(* CODESYS project RobotCell.project

Project tree, tasks and I/O mapping:
  Device : CODESYS Control Win V3 x64, CODESYS, version 3.5.22.40
    application Application
      libraries: Standard, 3.5.22.0 (System); VisuDialogs, * (System)
      task SoftMotion_PlanningTask (freewheeling, priority 15) calls nothing
      task CommTask (cyclic, interval t#50ms, priority 10) calls PRG_Comm
      task MainTask (cyclic, interval 4 ms, priority 1) calls PRG_Main, PRG_Tests, PRG_Recipe_Cell
      task VISU_TASK (cyclic, interval 100 ms, priority 31) calls VisuElems.Visu_Prg, PRG_HMI_Alarms, PRG_HMI_Robot, PRG_HMI_Overview
      axis group AxisGroup_Robot: TRAFO.Kin_ArticulatedRobot_6DOF, axes Axis_J1, Axis_J2, Axis_J3, Axis_J4, Axis_J5, Axis_J6
      Config/
        global variables GVL_Constants
        global variables GVL_CellGeometry
        global variables GVL_Params
        global variables GVL_Config
        global variables GVL_AlarmDefs
      Types/
        data type E_PackMLState
        data type E_PackMLMode
        data type E_PackMLCommand
        data type E_AlarmClass
        data type E_AlarmId
        data type E_Bin
        data type E_Quality
        data type E_DecisionSource
        data type E_PartState
        data type ST_PartRecord
        data type ST_AlarmDef
        data type ST_Alarm
        data type ST_VisionMsg
        data type ST_DecisionMsg
        data type ST_CaptureMsg
        data type E_RobotCmd
        data type E_PickStep
      Interfaces/
        interface I_AlarmSink: Raise, Clear, RaiseEvent
        interface I_Equipment: Reset, HasError, ErrorId
      Framework/
        function block FB_PackMLStateMachine [ST]
        function block FB_AlarmHandler [ST]: Raise, Clear, AcknowledgeAll, GetAlarm, RaiseEvent
        function block FB_PartQueue [ST]: AddRecord, FindIndex, GetRecord, PutRecord, Release, Count, Clear
      Equipment/
        function block FB_PhotoEye [ST]
        function block FB_Bin [ST]: Empty
        function block FB_SafetyMonitor [ST]
        function block FB_VacuumGripper [ST]: Reset, HasError, ErrorId
        function block FB_Conveyor [ST]: Reset, HasError, ErrorId
        function block FB_Robot [ST]: Reset, HasError, ErrorId
        function block FB_JointMonitor [ST]
        function block FB_CameraTrigger [ST]
      Process/
        function F_SelectBin [ST]
        function block FB_PartTracker [ST]: Decide, RaiseAlarm, CurrentX, NextPickable, FindPart, GetRecord, SetState, Count, RaiseEventAlarm, Clear
        function block FB_PickSequence [ST]: Request, NextStep, TrackedPose, GoError
        function block FB_SortingCell [ST]: AlarmState, PlacedCount, RobotMoving, AnyBinFull
      Comm/
        global variables GVL_Bridge
        global variables GVL_Hmi
        function block FB_MessageIntake [ST]
        function block FB_BridgeWatchdog [ST]
      Programs/
        program PRG_Main [ST]
        program PRG_Comm [ST]
      Tests/
        program PRG_TestMotionSmoke [ST]
        program PRG_Tests [ST]
        program PRG_TestTypes [ST]
        program PRG_TestPackML [ST]
        program PRG_TestAlarms [ST]
        program PRG_TestEquipment [ST]
        program PRG_TestMotion [ST]
        program PRG_TestTracking [ST]
        program PRG_TestJointMonitor [ST]
        program PRG_TestPick [ST]
        program PRG_TestCell [ST]
      visualisation Visu_Overview
      data type ST_Recipe_Cell
      global variables GVL_Recipe_Cell
      program PRG_Recipe_Cell [ST]
      Hmi/
        global variables GVL_HmiPanel
        global variables GVL_HmiView
        function block FB_HmiPanel [ST]
        function block FB_HmiView [ST]
      program PRG_HMI_Alarms [ST]
      visualisation Visu_Robot
      image pool IP_Robot
      program PRG_HMI_Robot [ST]
      program PRG_HMI_Overview [ST]
      image pool IP_Overview
      visualisation Visu_Alarms
      image pool IP_Alarms
    SoftMotion General Axis Pool : SoftMotion General Axis Pool, CODESYS, version 4.11.0.0
      Axis_J1 : SM_Drive_Virtual, CODESYS, order no. 1805, version 4.18.0.0
          settings: wDriveID = 0; fSWMaxVelocity = 180; fSWLimitPositive = 170; fSWLimitNegative = -170; bSWLimitEnable = true
      Axis_J2 : SM_Drive_Virtual, CODESYS, order no. 1805, version 4.18.0.0
          settings: fSWMaxVelocity = 180; fSWLimitPositive = 150; fSWLimitNegative = -90; bSWLimitEnable = true
      Axis_J3 : SM_Drive_Virtual, CODESYS, order no. 1805, version 4.18.0.0
          settings: wDriveID = 2; fSWMaxVelocity = 180; fSWLimitPositive = 150; fSWLimitNegative = -120; bSWLimitEnable = true
      Axis_J4 : SM_Drive_Virtual, CODESYS, order no. 1805, version 4.18.0.0
          settings: wDriveID = 3; fSWMaxVelocity = 360; fSWLimitPositive = 180; fSWLimitNegative = -180; bSWLimitEnable = true
      Axis_J5 : SM_Drive_Virtual, CODESYS, order no. 1805, version 4.18.0.0
          settings: wDriveID = 4; fSWMaxVelocity = 360; fSWLimitPositive = 120; fSWLimitNegative = -120; bSWLimitEnable = true
      Axis_J6 : SM_Drive_Virtual, CODESYS, order no. 1805, version 4.18.0.0
          settings: wDriveID = 5; fSWMaxVelocity = 360; fSWLimitPositive = 360; fSWLimitNegative = -360; bSWLimitEnable = true
      Axis_Conveyor : SM_Drive_Virtual, CODESYS, order no. 1805, version 4.18.0.0
          settings: wDriveID = 6; fSWMaxVelocity = 400; bSWLimitEnable = false
  libraries: VisuSymbols, 4.5.0.0 (System)
  5ce3da45-db07-42e7-a21c-a00fff4ed8f6|C:\Users\AvazA\AppData\Local\Temp\cmcp-visu-UXzo4K\ic_alarm_24_80868c.svg
  5ce3da45-db07-42e7-a21c-a00fff4ed8f6|C:\Users\AvazA\AppData\Local\Temp\cmcp-visu-UXzo4K\ic_check_27_1a232d.svg
  5ce3da45-db07-42e7-a21c-a00fff4ed8f6|C:\Users\AvazA\AppData\Local\Temp\cmcp-visu-UXzo4K\ic_pause_27_1a232d.svg
  5ce3da45-db07-42e7-a21c-a00fff4ed8f6|C:\Users\AvazA\AppData\Local\Temp\cmcp-visu-UXzo4K\ic_play_27_1a232d.svg
  5ce3da45-db07-42e7-a21c-a00fff4ed8f6|C:\Users\AvazA\AppData\Local\Temp\cmcp-visu-UXzo4K\stn_bin_on_48x48.svg
  5ce3da45-db07-42e7-a21c-a00fff4ed8f6|C:\Users\AvazA\AppData\Local\Temp\cmcp-visu-vSJax5\ic_stop_30_66727e.svg
  5ce3da45-db07-42e7-a21c-a00fff4ed8f6|C:\Users\AvazA\AppData\Local\Temp\cmcp-visu-vSJax5\ic_fault_30_d72332.svg
  5ce3da45-db07-42e7-a21c-a00fff4ed8f6|C:\Users\AvazA\AppData\Local\Temp\cmcp-visu-vSJax5\ic_pause_30_ffbb00.svg
  5ce3da45-db07-42e7-a21c-a00fff4ed8f6|C:\Users\AvazA\AppData\Local\Temp\cmcp-visu-vSJax5\ic_warning_30_ffbb00.svg
  5ce3da45-db07-42e7-a21c-a00fff4ed8f6|C:\Users\AvazA\AppData\Local\Temp\cmcp-visu-vSJax5\ic_manual_30_2f5d8a.svg
  5ce3da45-db07-42e7-a21c-a00fff4ed8f6|C:\Users\AvazA\AppData\Local\Temp\cmcp-visu-vSJax5\ic_play_30_66727e.svg
  5ce3da45-db07-42e7-a21c-a00fff4ed8f6|C:\Users\AvazA\AppData\Local\Temp\cmcp-visu-vSJax5\ic_login_27_1a232d.svg
  5ce3da45-db07-42e7-a21c-a00fff4ed8f6|C:\Users\AvazA\AppData\Local\Temp\cmcp-visu-vSJax5\ic_reset_27_1a232d.svg
  5ce3da45-db07-42e7-a21c-a00fff4ed8f6|C:\Users\AvazA\AppData\Local\Temp\cmcp-visu-vSJax5\ic_play_27_ffffff.svg
  5ce3da45-db07-42e7-a21c-a00fff4ed8f6|C:\Users\AvazA\AppData\Local\Temp\cmcp-visu-UXzo4K\sign_warning_30.svg
  5ce3da45-db07-42e7-a21c-a00fff4ed8f6|C:\Users\AvazA\AppData\Local\Temp\cmcp-visu-UXzo4K\ic_speed_24_80868c.svg
  5ce3da45-db07-42e7-a21c-a00fff4ed8f6|C:\Users\AvazA\AppData\Local\Temp\cmcp-visu-UXzo4K\ic_warning_30_ffbb00.svg
  5ce3da45-db07-42e7-a21c-a00fff4ed8f6|C:\Users\AvazA\AppData\Local\Temp\cmcp-visu-UXzo4K\ic_pause_30_ffbb00.svg
  5ce3da45-db07-42e7-a21c-a00fff4ed8f6|C:\Users\AvazA\AppData\Local\Temp\cmcp-visu-UXzo4K\ic_fault_30_d72332.svg
  5ce3da45-db07-42e7-a21c-a00fff4ed8f6|C:\Users\AvazA\AppData\Local\Temp\cmcp-visu-UXzo4K\ic_count_24_80868c.svg
  5ce3da45-db07-42e7-a21c-a00fff4ed8f6|C:\Users\AvazA\AppData\Local\Temp\cmcp-visu-UXzo4K\stn_bin_off_48x48.svg
  text list GlobalTextList
  5ce3da45-db07-42e7-a21c-a00fff4ed8f6|C:\Users\AvazA\AppData\Local\Temp\cmcp-visu-vSJax5\ic_stop_27_1a232d.svg
  5ce3da45-db07-42e7-a21c-a00fff4ed8f6|C:\Users\AvazA\AppData\Local\Temp\cmcp-visu-vSJax5\ic_home_33_5c636a.svg
  5ce3da45-db07-42e7-a21c-a00fff4ed8f6|C:\Users\AvazA\AppData\Local\Temp\cmcp-visu-vSJax5\ic_machine_33_2f5d8a.svg
  5ce3da45-db07-42e7-a21c-a00fff4ed8f6|C:\Users\AvazA\AppData\Local\Temp\cmcp-visu-vSJax5\ic_alarm_33_5c636a.svg
  5ce3da45-db07-42e7-a21c-a00fff4ed8f6|C:\Users\AvazA\AppData\Local\Temp\cmcp-visu-vSJax5\ic_manual_24_80868c.svg
  5ce3da45-db07-42e7-a21c-a00fff4ed8f6|C:\Users\AvazA\AppData\Local\Temp\cmcp-visu-vSJax5\ic_info_24_80868c.svg
  5ce3da45-db07-42e7-a21c-a00fff4ed8f6|C:\Users\AvazA\AppData\Local\Temp\cmcp-visu-vSJax5\ic_speed_24_80868c.svg
  5ce3da45-db07-42e7-a21c-a00fff4ed8f6|C:\Users\AvazA\AppData\Local\Temp\cmcp-visu-vSJax5\ic_machine_24_80868c.svg
  5ce3da45-db07-42e7-a21c-a00fff4ed8f6|C:\Users\AvazA\AppData\Local\Temp\cmcp-visu-UXzo4K\stn_robot6_off_48x48.svg
  5ce3da45-db07-42e7-a21c-a00fff4ed8f6|C:\Users\AvazA\AppData\Local\Temp\cmcp-visu-UXzo4K\ic_manual_23_2f5d8a.svg
  5ce3da45-db07-42e7-a21c-a00fff4ed8f6|C:\Users\AvazA\AppData\Local\Temp\cmcp-visu-UXzo4K\stn_camera_on_48x48.svg
  5ce3da45-db07-42e7-a21c-a00fff4ed8f6|C:\Users\AvazA\AppData\Local\Temp\cmcp-visu-UXzo4K\stn_camera_off_48x48.svg
  5ce3da45-db07-42e7-a21c-a00fff4ed8f6|C:\Users\AvazA\AppData\Local\Temp\cmcp-visu-UXzo4K\sign_alarm_27.svg
  5ce3da45-db07-42e7-a21c-a00fff4ed8f6|C:\Users\AvazA\AppData\Local\Temp\cmcp-visu-UXzo4K\stn_conveyor_on_48x14.svg
  5ce3da45-db07-42e7-a21c-a00fff4ed8f6|C:\Users\AvazA\AppData\Local\Temp\cmcp-visu-UXzo4K\stn_conveyor_off_48x14.svg
  5ce3da45-db07-42e7-a21c-a00fff4ed8f6|C:\Users\AvazA\AppData\Local\Temp\cmcp-visu-UXzo4K\sign_stop_13.svg
  5ce3da45-db07-42e7-a21c-a00fff4ed8f6|C:\Users\AvazA\AppData\Local\Temp\cmcp-visu-UXzo4K\sign_run_15.svg
  5ce3da45-db07-42e7-a21c-a00fff4ed8f6|C:\Users\AvazA\AppData\Local\Temp\cmcp-visu-UXzo4K\arrow_r_15_92979b.svg
  5ce3da45-db07-42e7-a21c-a00fff4ed8f6|C:\Users\AvazA\AppData\Local\Temp\cmcp-visu-UXzo4K\ic_alarm_33_5c636a.svg
  5ce3da45-db07-42e7-a21c-a00fff4ed8f6|C:\Users\AvazA\AppData\Local\Temp\cmcp-visu-UXzo4K\ic_machine_33_5c636a.svg
  5ce3da45-db07-42e7-a21c-a00fff4ed8f6|C:\Users\AvazA\AppData\Local\Temp\cmcp-visu-UXzo4K\ic_home_33_2f5d8a.svg
  5ce3da45-db07-42e7-a21c-a00fff4ed8f6|C:\Users\AvazA\AppData\Local\Temp\cmcp-visu-UXzo4K\ic_stop_27_1a232d.svg
  5ce3da45-db07-42e7-a21c-a00fff4ed8f6|C:\Users\AvazA\AppData\Local\Temp\cmcp-visu-UXzo4K\ic_play_27_ffffff.svg
  5ce3da45-db07-42e7-a21c-a00fff4ed8f6|C:\Users\AvazA\AppData\Local\Temp\cmcp-visu-UXzo4K\ic_reset_27_1a232d.svg
  5ce3da45-db07-42e7-a21c-a00fff4ed8f6|C:\Users\AvazA\AppData\Local\Temp\cmcp-visu-UXzo4K\ic_login_27_1a232d.svg
  5ce3da45-db07-42e7-a21c-a00fff4ed8f6|C:\Users\AvazA\AppData\Local\Temp\cmcp-visu-UXzo4K\ic_play_30_66727e.svg
  5ce3da45-db07-42e7-a21c-a00fff4ed8f6|C:\Users\AvazA\AppData\Local\Temp\cmcp-visu-UXzo4K\ic_manual_30_2f5d8a.svg
  5ce3da45-db07-42e7-a21c-a00fff4ed8f6|C:\Users\AvazA\AppData\Local\Temp\cmcp-visu-UXzo4K\ic_stop_30_66727e.svg
  5ce3da45-db07-42e7-a21c-a00fff4ed8f6|C:\Users\AvazA\AppData\Local\Temp\cmcp-visu-UXzo4K\stn_robot6_on_48x48.svg
  5ce3da45-db07-42e7-a21c-a00fff4ed8f6|C:\Users\AvazA\AppData\Local\Temp\cmcp-visu-UXzo4K\stn_gripper_on_48x48.svg
  5ce3da45-db07-42e7-a21c-a00fff4ed8f6|C:\Users\AvazA\AppData\Local\Temp\cmcp-visu-UXzo4K\stn_gripper_off_48x48.svg
  5ce3da45-db07-42e7-a21c-a00fff4ed8f6|C:\Users\AvazA\AppData\Local\Temp\cmcp-visu-6UqmBO\ic_check_27_1a232d.svg
  5ce3da45-db07-42e7-a21c-a00fff4ed8f6|C:\Users\AvazA\AppData\Local\Temp\cmcp-visu-6UqmBO\ic_warning_24_80868c.svg
  5ce3da45-db07-42e7-a21c-a00fff4ed8f6|C:\Users\AvazA\AppData\Local\Temp\cmcp-visu-6UqmBO\ic_alarm_24_80868c.svg
  5ce3da45-db07-42e7-a21c-a00fff4ed8f6|C:\Users\AvazA\AppData\Local\Temp\cmcp-visu-6UqmBO\ic_alarm_33_2f5d8a.svg
  5ce3da45-db07-42e7-a21c-a00fff4ed8f6|C:\Users\AvazA\AppData\Local\Temp\cmcp-visu-6UqmBO\ic_machine_33_5c636a.svg
  5ce3da45-db07-42e7-a21c-a00fff4ed8f6|C:\Users\AvazA\AppData\Local\Temp\cmcp-visu-6UqmBO\ic_home_33_5c636a.svg
  5ce3da45-db07-42e7-a21c-a00fff4ed8f6|C:\Users\AvazA\AppData\Local\Temp\cmcp-visu-6UqmBO\ic_stop_27_1a232d.svg
  5ce3da45-db07-42e7-a21c-a00fff4ed8f6|C:\Users\AvazA\AppData\Local\Temp\cmcp-visu-6UqmBO\ic_play_27_ffffff.svg
  5ce3da45-db07-42e7-a21c-a00fff4ed8f6|C:\Users\AvazA\AppData\Local\Temp\cmcp-visu-6UqmBO\ic_reset_27_1a232d.svg
  5ce3da45-db07-42e7-a21c-a00fff4ed8f6|C:\Users\AvazA\AppData\Local\Temp\cmcp-visu-6UqmBO\ic_login_27_1a232d.svg
  5ce3da45-db07-42e7-a21c-a00fff4ed8f6|C:\Users\AvazA\AppData\Local\Temp\cmcp-visu-6UqmBO\ic_play_30_66727e.svg
  5ce3da45-db07-42e7-a21c-a00fff4ed8f6|C:\Users\AvazA\AppData\Local\Temp\cmcp-visu-6UqmBO\ic_manual_30_2f5d8a.svg
  5ce3da45-db07-42e7-a21c-a00fff4ed8f6|C:\Users\AvazA\AppData\Local\Temp\cmcp-visu-6UqmBO\ic_warning_30_ffbb00.svg
  5ce3da45-db07-42e7-a21c-a00fff4ed8f6|C:\Users\AvazA\AppData\Local\Temp\cmcp-visu-6UqmBO\ic_pause_30_ffbb00.svg
  5ce3da45-db07-42e7-a21c-a00fff4ed8f6|C:\Users\AvazA\AppData\Local\Temp\cmcp-visu-6UqmBO\ic_fault_30_d72332.svg
  5ce3da45-db07-42e7-a21c-a00fff4ed8f6|C:\Users\AvazA\AppData\Local\Temp\cmcp-visu-6UqmBO\ic_stop_30_66727e.svg
  5ce3da45-db07-42e7-a21c-a00fff4ed8f6|C:\Users\AvazA\AppData\Local\Temp\cmcp-visu-UXzo4K\ic_info_24_80868c.svg
*)

// Device/Application/Types/E_PackMLState
// PackML unit states, numbered as in ISA-TR88.00.02.
{attribute 'qualified_only'}
{attribute 'strict'}
TYPE E_PackMLState :
(
    Undefined := 0,
    Clearing := 1,
    Stopped := 2,
    Starting := 3,
    Idle := 4,
    Suspended := 5,
    Execute := 6,
    Stopping := 7,
    Aborting := 8,
    Aborted := 9,
    Holding := 10,
    Held := 11,
    Unholding := 12,
    Suspending := 13,
    Unsuspending := 14,
    Resetting := 15,
    Completing := 16,
    Complete := 17
);
END_TYPE

// Device/Application/Types/E_PackMLMode
// PackML unit modes used by this cell.
{attribute 'qualified_only'}
{attribute 'strict'}
TYPE E_PackMLMode :
(
    Production := 1,
    Maintenance := 2,
    Manual := 3
);
END_TYPE

// Device/Application/Types/E_PackMLCommand
// PackML state commands.
{attribute 'qualified_only'}
{attribute 'strict'}
TYPE E_PackMLCommand :
(
    None := 0,
    Reset := 1,
    Start := 2,
    Stop := 3,
    Hold := 4,
    Unhold := 5,
    Suspend := 6,
    Unsuspend := 7,
    Abort := 8,
    Clear := 9,
    Complete := 10
);
END_TYPE

// Device/Application/Types/E_AlarmClass
// Alarm classes (ISA-18.2 style priorities). Critical -> Abort, Error -> Stop.
{attribute 'qualified_only'}
{attribute 'strict'}
TYPE E_AlarmClass :
(
    Info := 0,
    Warning := 1,
    Error := 2,
    Critical := 3
);
END_TYPE

// Device/Application/Types/E_AlarmId
// Every alarm of the cell. Definitions (class, text) are in GVL_AlarmDefs.
{attribute 'qualified_only'}
{attribute 'strict'}
TYPE E_AlarmId :
(
    None := 0,
    EStop := 1,
    DoorOpen := 2,
    BridgeLost := 3,
    AxisGroupError := 4,
    ConveyorError := 5,
    FollowingErrorWarn := 6,
    FollowingErrorFault := 7,
    FeedbackStale := 8,
    VacuumNoGrip := 9,
    VacuumLost := 10,
    PartMissed := 11,
    BinFull := 12,
    VisionMissing := 13,
    DecisionFallback := 14,
    LowConfidence := 15,
    QueueOverflow := 16
);
END_TYPE

// Device/Application/Types/E_Bin
// Output bins: one per good part type, then the quality bins.
{attribute 'qualified_only'}
{attribute 'strict'}
TYPE E_Bin :
(
    TypeA := 0,
    TypeB := 1,
    TypeC := 2,
    Rework := 3,
    Scrap := 4,
    Quarantine := 5
);
END_TYPE

// Device/Application/Types/E_Quality
// Quality disposition of a part (spec section 6.3).
{attribute 'qualified_only'}
{attribute 'strict'}
TYPE E_Quality :
(
    Unknown := 0,
    Ok := 1,
    Rework := 2,
    Scrap := 3
);
END_TYPE

// Device/Application/Types/E_DecisionSource
// Where a part's quality decision came from.
{attribute 'qualified_only'}
{attribute 'strict'}
TYPE E_DecisionSource :
(
    None := 0,
    Ai := 1,
    Fallback := 2
);
END_TYPE

// Device/Application/Types/E_PartState
// Life cycle of a tracked part.
{attribute 'qualified_only'}
{attribute 'strict'}
TYPE E_PartState :
(
    Free := 0,
    Captured := 1,
    Identified := 2,
    Decided := 3,
    Scheduled := 4,
    Picked := 5,
    Placed := 6,
    Missed := 7,
    Dropped := 8
);
END_TYPE

// Device/Application/Types/ST_PartRecord
// One tracked part. Positions are in the belt frame at capture time (mm, degrees).
TYPE ST_PartRecord :
STRUCT
    udiPartId : UDINT;
    lrBeltPosAtCapture : LREAL;         // conveyor axis position when PE1 triggered [mm]
    xVisionValid : BOOL;
    usiClass : USINT;                   // detector class index 0..2
    rConfidence : REAL;                 // detector confidence 0..1
    lrX : LREAL;                        // belt frame X at capture [mm]
    lrY : LREAL;                        // belt frame Y [mm]
    lrTheta : LREAL;                    // orientation about Z [deg]
    eQuality : E_Quality;
    rQualityProb : REAL;                // probability of the chosen quality option
    xIdentReliable : BOOL;
    eDecisionSource : E_DecisionSource;
    eTargetBin : E_Bin;
    eState : E_PartState;
    tCaptured : TIME;                   // TIME() at capture
END_STRUCT
END_TYPE

// Device/Application/Types/ST_AlarmDef
// Static definition of one alarm.
TYPE ST_AlarmDef :
STRUCT
    eClass : E_AlarmClass;
    sText : STRING(80);
END_STRUCT
END_TYPE

// Device/Application/Types/ST_Alarm
// Runtime state of one alarm.
TYPE ST_Alarm :
STRUCT
    eClass : E_AlarmClass;
    xActive : BOOL;
    xAcked : BOOL := TRUE;              // no pending acknowledgement
    tRaised : TIME;
END_STRUCT
END_TYPE

// Device/Application/Types/ST_VisionMsg
// Vision result written by the bridge. A new message has a new udiSeq.
TYPE ST_VisionMsg :
STRUCT
    udiSeq : UDINT;
    udiPartId : UDINT;
    xValid : BOOL;
    usiClass : USINT;
    rConfidence : REAL;
    lrX : LREAL;                        // belt frame [mm]
    lrY : LREAL;                        // belt frame [mm]
    lrTheta : LREAL;                    // [deg]
END_STRUCT
END_TYPE

// Device/Application/Types/ST_DecisionMsg
// Quality decision written by the bridge (THX-02). A new message has a new udiSeq.
TYPE ST_DecisionMsg :
STRUCT
    udiSeq : UDINT;
    udiPartId : UDINT;
    eQuality : E_Quality;
    rQualityProb : REAL;
    xIdentReliable : BOOL;
END_STRUCT
END_TYPE

// Device/Application/Types/ST_CaptureMsg
// Capture request from the PLC to the bridge. A new request has a new udiSeq.
TYPE ST_CaptureMsg :
STRUCT
    udiSeq : UDINT;
    udiPartId : UDINT;
    lrBeltPos : LREAL;                  // conveyor axis position at the trigger [mm]
END_STRUCT
END_TYPE

// Device/Application/Types/E_RobotCmd
// Commands of FB_Robot (start on a rising edge of xExecute).
{attribute 'qualified_only'}
{attribute 'strict'}
TYPE E_RobotCmd :
(
    None := 0,
    MovePtpAcs := 1,       // point-to-point, target in joint space
    MoveLinMcs := 2,       // linear, target in machine coordinates
    MoveLinPcs1 := 3,      // linear, target in PCS_1 (conveyor tracking frame)
    Stop := 4,             // controlled stop, aborts any motion
    Reset := 5,            // reset axis group errors
    MovePtpMcs := 6        // point-to-point, Cartesian target in machine coordinates
);
END_TYPE

// Device/Application/Types/E_PickStep
// Steps of FB_PickSequence.
{attribute 'qualified_only'}
{attribute 'strict'}
TYPE E_PickStep :
(
    Idle := 0,
    MoveHome := 1,
    MoveReady := 2,
    WaitPart := 3,
    StartTracking := 4,
    Approach := 5,
    Descend := 6,
    Grip := 7,
    Lift := 8,
    MoveToBin := 9,
    Release := 10,
    Retract := 11,
    Aborting := 12,
    Aborted := 13,
    Error := 14,
    RecoverLift := 15       // after an abort with a part on the cup: straight up first
);
END_TYPE

// Device/Application/ST_Recipe_Cell
TYPE ST_Recipe_Cell :
STRUCT
    lrBeltSpeed : LREAL; // GVL_Params.lrBeltSpeed
    lrApproachHeight : LREAL; // GVL_Params.lrApproachHeight
    lrPickDepth : LREAL; // GVL_Params.lrPickDepth
    lrLinVelocity : LREAL; // GVL_Params.lrLinVelocity
    lrLinAccel : LREAL; // GVL_Params.lrLinAccel
    lrLinJerk : LREAL; // GVL_Params.lrLinJerk
    lrPtpVelFactor : LREAL; // GVL_Params.lrPtpVelFactor
    rConfidenceThreshold : REAL; // GVL_Params.rConfidenceThreshold
    tDecisionDeadline : TIME; // GVL_Params.tDecisionDeadline
    tVacuumTimeout : TIME; // GVL_Params.tVacuumTimeout
    lrFollowErrWarn : LREAL; // GVL_Params.lrFollowErrWarn
    lrFollowErrFault : LREAL; // GVL_Params.lrFollowErrFault
    tFeedbackTimeout : TIME; // GVL_Params.tFeedbackTimeout
END_STRUCT
END_TYPE

// Device/Application/Config/GVL_Constants
// Project-wide constants. Values that change per recipe live in GVL_Params, not here.
{attribute 'qualified_only'}
VAR_GLOBAL CONSTANT
    PROJECT_VERSION : STRING := '0.7.0';
END_VAR

// Device/Application/Config/GVL_CellGeometry
// Fixed geometry of the cell. Units: mm and degrees, robot base frame (Z up).
// Kinematics values must match the axis group AxisGroup_Robot (plc/scripts/build_softmotion_base.py).
// Orientations (A, B, C): B = 180 points the tool straight down (verified in simulation).
{attribute 'qualified_only'}
VAR_GLOBAL CONSTANT
    // Kin_ArticulatedRobot_6DOF parameters [mm]
    ROBOT_A1 : LREAL := 50;
    ROBOT_D1 : LREAL := 400;
    ROBOT_A2 : LREAL := 450;
    ROBOT_A3 : LREAL := 50;
    ROBOT_D3 : LREAL := 0;
    ROBOT_D4 : LREAL := 450;
    ROBOT_D6 : LREAL := 120;                 // flange + suction tool

    // Tool pointing straight down
    TOOL_DOWN_A : LREAL := 0;
    TOOL_DOWN_B : LREAL := 180;
    TOOL_DOWN_C : LREAL := 180;

    // Conveyor belt frame: origin at the infeed, +X along the flow direction.
    BELT_ORIGIN : MC_COORD_REF := (X := -1500, Y := -550, Z := 0, A := 0, B := 0, C := 0);
    BELT_SURFACE_Z : LREAL := 0;
    PE1_X : LREAL := 300;                    // camera trigger photo-eye, belt frame [mm]
    PE2_X : LREAL := 1050;                   // pick window start, belt frame [mm]
    PICK_WINDOW_END_X : LREAL := 1750;       // pick window end, belt frame [mm]
    PICK_MARGIN : LREAL := 300;              // do not start a pick this close to the window end [mm]
    // Grip height of each part class above the belt [mm]: the top surface under the suction
    // cup (config/parts.yaml classes, tools/fetch_objects.py meta.json; a unit test keeps
    // both equal)
    PART_HEIGHTS : ARRAY[0..2] OF LREAL := [56.39, 81.19, 83.46];

    // Home position, joint space [deg]
    HOME_ACS : SMC_POS_REF := (a := (a0 := 0, a1 := -30, a2 := 60, a3 := 0, a4 := 60, a5 := 0));
    // Waiting pose above the pick window, tool down (machine coordinates)
    READY_POSE : MC_COORD_REF := (X := -100, Y := -550, Z := 300, A := 0, B := 180, C := 180);
    RETRACT_HEIGHT : LREAL := 100;           // lift above the bin drop pose after release [mm]

    // Drop poses above the bins (tool pointing down), machine coordinates [mm, deg]. Z 300: a
    // held part up to 90 mm tall clears the 160 mm bin rim by 50 mm.
    BIN_DROP : ARRAY[E_Bin.TypeA..E_Bin.Quarantine] OF MC_COORD_REF := [
        (X := -500, Y := 550, Z := 300, A := 0, B := 180, C := 180),
        (X := -300, Y := 550, Z := 300, A := 0, B := 180, C := 180),
        (X := -100, Y := 550, Z := 300, A := 0, B := 180, C := 180),
        (X := 100, Y := 550, Z := 300, A := 0, B := 180, C := 180),
        (X := 300, Y := 550, Z := 300, A := 0, B := 180, C := 180),
        (X := 500, Y := 550, Z := 300, A := 0, B := 180, C := 180)];
END_VAR

// Device/Application/Config/GVL_Params
// Process parameters. Retained; written by the recipes (Standard / HighSpeed).
{attribute 'qualified_only'}
VAR_GLOBAL RETAIN
    lrBeltSpeed : LREAL := 100;              // conveyor speed [mm/s]
    lrApproachHeight : LREAL := 80;          // approach / lift height above the part [mm]
    lrPickDepth : LREAL := 5;                // how far below the part top the cup goes [mm]
    lrLinVelocity : LREAL := 500;            // linear path velocity [mm/s]
    lrLinAccel : LREAL := 2000;              // linear path acceleration [mm/s2]
    lrLinJerk : LREAL := 20000;              // linear path jerk [mm/s3]
    lrPtpVelFactor : LREAL := 0.5;           // PTP velocity factor ]0, 1]
    rConfidenceThreshold : REAL := 0.6;      // below this the part goes to quarantine
    tDecisionDeadline : TIME := T#2S500MS;   // fallback if no decision by then
    tVacuumTimeout : TIME := T#500MS;        // no grip -> error
    lrFollowErrWarn : LREAL := 2.0;          // following error warning [deg]
    lrFollowErrFault : LREAL := 5.0;         // following error fault [deg]
    tFeedbackTimeout : TIME := T#500MS;      // joint feedback must update within this time
    aClassToBin : ARRAY[0..2] OF E_Bin := [E_Bin.TypeA, E_Bin.TypeB, E_Bin.TypeC];
END_VAR

// Device/Application/Config/GVL_Config
// Build/run configuration.
{attribute 'qualified_only'}
VAR_GLOBAL
    // Joint feedback := setpoint (no staleness check) unless the twin reports itself active through
    // GVL_Bridge.xTwinActive. FALSE forces real feedback even without the twin.
    xFeedbackLoopback : BOOL := TRUE;
    // The sorting cell runs in PRG_Main. Simulation tests of single blocks switch it off so their
    // harnesses can own the robot and the conveyor.
    xCellEnabled : BOOL := TRUE;
END_VAR
VAR_GLOBAL CONSTANT
    MAX_PARTS : UINT := 32;                  // capacity of the part queue
END_VAR

// Device/Application/Config/GVL_AlarmDefs
// Alarm definitions: class and operator text for every E_AlarmId.
// Critical -> PackML Abort, Error -> Stop, Warning -> no state change (BinFull suspends the unit).
{attribute 'qualified_only'}
VAR_GLOBAL CONSTANT
    aDefs : ARRAY[E_AlarmId.None..E_AlarmId.QueueOverflow] OF ST_AlarmDef := [
        (eClass := E_AlarmClass.Info, sText := 'No alarm'),
        (eClass := E_AlarmClass.Critical, sText := 'Emergency stop pressed'),
        (eClass := E_AlarmClass.Critical, sText := 'Safety door opened in automatic mode'),
        (eClass := E_AlarmClass.Critical, sText := 'Connection to the digital twin bridge lost'),
        (eClass := E_AlarmClass.Critical, sText := 'Robot axis group error'),
        (eClass := E_AlarmClass.Error, sText := 'Conveyor axis error'),
        (eClass := E_AlarmClass.Warning, sText := 'Joint following error above warning limit'),
        (eClass := E_AlarmClass.Critical, sText := 'Joint following error above fault limit'),
        (eClass := E_AlarmClass.Critical, sText := 'Joint feedback not updated'),
        (eClass := E_AlarmClass.Error, sText := 'Vacuum not reached - part not gripped'),
        (eClass := E_AlarmClass.Error, sText := 'Vacuum lost while carrying a part'),
        (eClass := E_AlarmClass.Warning, sText := 'Part left the pick window unpicked'),
        (eClass := E_AlarmClass.Warning, sText := 'A bin is full - cell suspended until it is emptied'),
        (eClass := E_AlarmClass.Warning, sText := 'No vision result for a captured part'),
        (eClass := E_AlarmClass.Warning, sText := 'AI decision late - fallback rule used'),
        (eClass := E_AlarmClass.Warning, sText := 'Low detection confidence - part quarantined'),
        (eClass := E_AlarmClass.Error, sText := 'Part queue full')];
END_VAR

// Device/Application/Comm/GVL_Bridge
// Exchange with the Python bridge over OPC UA (published by the symbol configuration).
// Tag names for the bridge: config/opcua_tags.yaml. In Phase 1, tests write the inputs.
{attribute 'qualified_only'}
{attribute 'symbol' := 'readwrite'}
VAR_GLOBAL
    // --- inputs (bridge -> PLC) ---
    xHeartbeat : BOOL;                                     // toggled by the bridge every cycle
    xTwinActive : BOOL;                                    // the twin delivers joint feedback
    aJointPosFb : ARRAY[1..6] OF LREAL;                    // measured joint positions [deg]
    aJointTorqueFb : ARRAY[1..6] OF LREAL;                 // measured joint torques [Nm]
    udiFeedbackSeq : UDINT;                                // increments with every feedback sample
    udiFeedbackForSeq : UDINT;                             // udiSetpointSeq the feedback belongs to
    xPE1 : BOOL;                                           // photo-eye at the camera
    xPE2 : BOOL;                                           // photo-eye at the pick window start
    xVacuumOk : BOOL;                                      // vacuum switch of the suction cup
    axBinFull : ARRAY[E_Bin.TypeA..E_Bin.Quarantine] OF BOOL;
    xDoorClosed : BOOL := TRUE;                            // safety door (TRUE = closed)
    xEStopOk : BOOL := TRUE;                               // emergency stop circuit (TRUE = not pressed)
    stVision : ST_VisionMsg;
    stDecision : ST_DecisionMsg;
    xDecisionActive : BOOL;                                // an AI decision service answers stDecision
    // --- outputs (PLC -> bridge) ---
    aJointPosSp : ARRAY[1..6] OF LREAL;                    // joint setpoints [deg]
    udiSetpointSeq : UDINT;                                // increments with every setpoint sample
    lrBeltPos : LREAL;                                     // conveyor position [mm]
    lrBeltVel : LREAL;                                     // conveyor velocity [mm/s]
    xVacuumOn : BOOL;                                      // vacuum valve
    stCapture : ST_CaptureMsg;
    eState : E_PackMLState;
    eMode : E_PackMLMode;
    // --- diagnostics (PLC -> bridge, HMI) ---
    eNewestAlarm : E_AlarmId;
    xAlarmError : BOOL;                                    // an Error-class alarm is active
    xAlarmCritical : BOOL;                                 // a Critical-class alarm is active
    ePickStep : E_PickStep;
    iWorstJoint : INT;                                     // joint with the largest following error
    aFollowingError : ARRAY[1..6] OF LREAL;                // [deg]
END_VAR

// Device/Application/Comm/GVL_Hmi
// Operator commands from the HMI (CODESYS Visualization) and, for tests and the HMI of later
// phases, over OPC UA (published by the symbol configuration).
{attribute 'qualified_only'}
{attribute 'symbol' := 'readwrite'}
VAR_GLOBAL
    eCommand : E_PackMLCommand;
    eModeRequest : E_PackMLMode := E_PackMLMode.Production;
    xAlarmAck : BOOL;
    axJogPlus : ARRAY[1..6] OF BOOL;
    axJogMinus : ARRAY[1..6] OF BOOL;
    rOverride : REAL := 1.0;                               // speed override ]0, 1]
END_VAR

// Device/Application/GVL_Recipe_Cell
// Recipes 'Cell', generated by codesys-mcp-toolkit (create_recipes). RETAIN: values saved from the HMI survive a power cycle.
VAR_GLOBAL RETAIN
    aRecipes : ARRAY[0..1] OF ST_Recipe_Cell := [(lrBeltSpeed := 100.0, lrApproachHeight := 80.0, lrPickDepth := 5.0, lrLinVelocity := 500.0, lrLinAccel := 2000.0, lrLinJerk := 20000.0, lrPtpVelFactor := 0.5, rConfidenceThreshold := 0.6, tDecisionDeadline := T#2S500MS, tVacuumTimeout := T#500MS, lrFollowErrWarn := 2.0, lrFollowErrFault := 5.0, tFeedbackTimeout := T#500MS), (lrBeltSpeed := 200.0, lrApproachHeight := 80.0, lrPickDepth := 5.0, lrLinVelocity := 800.0, lrLinAccel := 3000.0, lrLinJerk := 20000.0, lrPtpVelFactor := 0.8, rConfidenceThreshold := 0.6, tDecisionDeadline := T#2S500MS, tVacuumTimeout := T#500MS, lrFollowErrWarn := 2.0, lrFollowErrFault := 5.0, tFeedbackTimeout := T#500MS)];
END_VAR
VAR_GLOBAL CONSTANT
    asNames : ARRAY[0..1] OF STRING(32) := ['Standard', 'HighSpeed'];
    iCount : INT := 2;
END_VAR

// Device/Application/Hmi/GVL_HmiPanel
// Operator panel of the CODESYS Visualization: buttons and selectors write here; FB_HmiPanel
// turns them into the cell's commands (GVL_Hmi). Buttons are one-shot: cleared after use.
{attribute 'qualified_only'}
VAR_GLOBAL
    xStart : BOOL;
    xStop : BOOL;
    xReset : BOOL;
    xClear : BOOL;
    xAbort : BOOL;
    xSuspend : BOOL;
    xUnsuspend : BOOL;
    xAckAll : BOOL;                                        // acknowledge all alarms
    iModeSelect : INT := 1;                                // 1 Production, 2 Maintenance, 3 Manual
END_VAR

// Device/Application/Hmi/GVL_HmiView
// Display data for the CODESYS Visualization, prepared by FB_HmiView (no logic in screens).
{attribute 'qualified_only'}
VAR_GLOBAL
    sState : STRING(20);                                   // PackML state
    sMode : STRING(20);                                    // PackML mode
    sPickStep : STRING(20);                                // robot sequence step
    sNewestAlarm : STRING(80);                             // text of the newest alarm
    xExecute : BOOL;                                       // state groups for the machine bar
    xStopped : BOOL;
    xIdle : BOOL;
    xAborted : BOOL;                                       // Aborting or Aborted
    xHeld : BOOL;                                          // Held, Suspended or their acting states
    xActing : BOOL;                                        // Resetting, Starting, Stopping, Clearing
    xManual : BOOL;
    xAnyAlarm : BOOL;                                      // an alarm is active or unacknowledged
    axAlarm : ARRAY[1..16] OF BOOL;                        // per E_AlarmId: active or unacknowledged
    axAlarmActive : ARRAY[1..16] OF BOOL;                  // per E_AlarmId: condition present
    uiPlaced : UINT;                                       // parts placed (all bins)
    xBeltRunning : BOOL;                                   // conveyor faster than BELT_RUNNING_MM_S
    xRobotMoving : BOOL;                                   // a robot motion command is active
    xAnyBinFull : BOOL;                                    // at least one bin reports full
    xJogPermitted : BOOL;                                  // Manual mode and Execute: jog buttons act
END_VAR

// Device/Application/Programs/PRG_Comm
(*
    PRG_Comm
    Purpose : Communication entry point: OPC UA data consistency and statistics (Phase 2).
    Task    : CommTask, cyclic 50 ms
    Rule    : thin program - only instantiation and calls, no logic.
*)
PROGRAM PRG_Comm
VAR
END_VAR

// Intentionally empty until Phase 2.

END_PROGRAM

// Device/Application/Programs/PRG_Main
(*
    PRG_Main
    Purpose : Cell entry point: maps the bridge and HMI variable lists to the sorting cell unit.
    Task    : MainTask, cyclic 4 ms, SoftMotion bus cycle task
    Rule    : thin program - only instantiation, mapping and calls, no logic.
    Commands: GVL_Hmi.eCommand / xAlarmAck are written asynchronously (HMI, OPC UA). They are
              read once per cycle into a snapshot and cleared only if they still hold that
              value, so a command written during the cycle is never lost.
    HMI     : fbHmiPanel turns the visualization's buttons into GVL_Hmi commands before the
              snapshot; fbHmiView prepares GVL_HmiView after the cell has run.
    OPC UA  : published read-only for diagnostics (alarms, pick step) and the HMI.
*)
PROGRAM PRG_Main
{attribute 'symbol' := 'read'}
VAR
    sProjectVersion : STRING := GVL_Constants.PROJECT_VERSION;  // diagnostics: project version visible online and via OPC UA
    fbCell : FB_SortingCell;
    fbHmiPanel : FB_HmiPanel;
    fbHmiView : FB_HmiView;
    eCommand : E_PackMLCommand;
    xAlarmAck : BOOL;
END_VAR

IF NOT GVL_Config.xCellEnabled THEN
    RETURN;
END_IF

fbHmiPanel();
eCommand := GVL_Hmi.eCommand;
xAlarmAck := GVL_Hmi.xAlarmAck;
fbCell(AxisGroup := AxisGroup_Robot,
       ConveyorAxis := Axis_Conveyor,
       eCommand := eCommand,
       eModeRequest := GVL_Hmi.eModeRequest,
       xAlarmAck := xAlarmAck,
       axJogPlus := GVL_Hmi.axJogPlus,
       axJogMinus := GVL_Hmi.axJogMinus,
       rOverride := GVL_Hmi.rOverride,
       xHeartbeat := GVL_Bridge.xHeartbeat,
       aJointPosFb := GVL_Bridge.aJointPosFb,
       aJointTorqueFb := GVL_Bridge.aJointTorqueFb,
       udiFeedbackSeq := GVL_Bridge.udiFeedbackSeq,
       udiFeedbackForSeq := GVL_Bridge.udiFeedbackForSeq,
       xPE1 := GVL_Bridge.xPE1,
       xVacuumOk := GVL_Bridge.xVacuumOk,
       axBinFull := GVL_Bridge.axBinFull,
       xDoorClosed := GVL_Bridge.xDoorClosed,
       xEStopOk := GVL_Bridge.xEStopOk,
       stVision := GVL_Bridge.stVision,
       stDecision := GVL_Bridge.stDecision,
       xDecisionActive := GVL_Bridge.xDecisionActive,
       // joint feedback from the twin once the bridge reports it active (ADR 0008)
       xLoopback := GVL_Config.xFeedbackLoopback AND NOT GVL_Bridge.xTwinActive,
       aJointPosSp => GVL_Bridge.aJointPosSp,
       udiSetpointSeq => GVL_Bridge.udiSetpointSeq,
       lrBeltPos => GVL_Bridge.lrBeltPos,
       lrBeltVel => GVL_Bridge.lrBeltVel,
       xVacuumOn => GVL_Bridge.xVacuumOn,
       stCapture => GVL_Bridge.stCapture,
       eState => GVL_Bridge.eState,
       eMode => GVL_Bridge.eMode,
       ePickStep => GVL_Bridge.ePickStep,
       eNewestAlarm => GVL_Bridge.eNewestAlarm,
       xAlarmError => GVL_Bridge.xAlarmError,
       xAlarmCritical => GVL_Bridge.xAlarmCritical,
       iWorstJoint => GVL_Bridge.iWorstJoint,
       aFollowingError => GVL_Bridge.aFollowingError);
// commands are one-shot: consume the value this cycle has seen, keep a newer one
IF GVL_Hmi.eCommand = eCommand THEN
    GVL_Hmi.eCommand := E_PackMLCommand.None;
END_IF
IF xAlarmAck THEN
    GVL_Hmi.xAlarmAck := FALSE;
END_IF
fbHmiView(Cell := fbCell);

END_PROGRAM

// Device/Application/Process/FB_SortingCell
(*
    FB_SortingCell
    Purpose : The sorting cell as one PackML unit. Owns all equipment and maps the PackML states
              to equipment actions; computes the interlocks.
    In/Out  : AxisGroup (AxisGroup_Robot), ConveyorAxis (Axis_Conveyor)
    Inputs  : operator commands (GVL_Hmi), sensors and messages (GVL_Bridge), xLoopback (feedback := setpoint)
    Outputs : setpoints, belt and vacuum to the bridge; eState, eMode, ePickStep, aActAcs;
              diagnostics (newest alarm, alarm classes, worst joint, following errors)
    States  : Resetting  - acknowledge alarms, reset equipment and the pick sequence, forget the
                           tracked parts; done when safe and fault-free
              Starting / Unholding / Unsuspending - robot home -> ready, conveyor at speed
                           (a part still on the cup is placed in quarantine first)
              Execute    - automatic: pick sequence runs; Manual: jogging
              Stopping / Holding / Suspending / Completing - finish the current part, go home;
                           done when the sequence rests, the robot and the belt stand still
              Aborting   - controlled stop, vacuum kept; Clearing - reset the sequence
    Interlocks: Critical alarm or not safe -> Abort; Error alarm -> Stop; any bin full -> Suspend,
              and Unsuspend automatically when that bin is emptied (not after an operator Suspend).
              Resetting and Clearing are not interrupted by the alarms they are clearing.
*)
FUNCTION_BLOCK FB_SortingCell
VAR_IN_OUT
    AxisGroup : AXIS_GROUP_REF_SM3;
    ConveyorAxis : AXIS_REF_SM3;
END_VAR
VAR_INPUT
    eCommand : E_PackMLCommand;
    eModeRequest : E_PackMLMode := E_PackMLMode.Production;
    xAlarmAck : BOOL;
    axJogPlus : ARRAY[1..6] OF BOOL;
    axJogMinus : ARRAY[1..6] OF BOOL;
    rOverride : REAL := 1.0;
    xHeartbeat : BOOL;
    aJointPosFb : ARRAY[1..6] OF LREAL;
    aJointTorqueFb : ARRAY[1..6] OF LREAL;
    udiFeedbackSeq : UDINT;
    udiFeedbackForSeq : UDINT;                // setpoint sample the joint feedback answers
    xPE1 : BOOL;
    xVacuumOk : BOOL;
    axBinFull : ARRAY[E_Bin.TypeA..E_Bin.Quarantine] OF BOOL;
    xDoorClosed : BOOL := TRUE;
    xEStopOk : BOOL := TRUE;
    stVision : ST_VisionMsg;
    stDecision : ST_DecisionMsg;
    xDecisionActive : BOOL;                  // an AI decision service answers (bridge)
    xLoopback : BOOL;
END_VAR
VAR_OUTPUT
    aJointPosSp : ARRAY[1..6] OF LREAL;
    lrBeltPos : LREAL;
    lrBeltVel : LREAL;
    xVacuumOn : BOOL;
    stCapture : ST_CaptureMsg;
    eState : E_PackMLState := E_PackMLState.Stopped;
    eMode : E_PackMLMode := E_PackMLMode.Production;
    ePickStep : E_PickStep;
    aActAcs : ARRAY[1..6] OF LREAL;
    udiSetpointSeq : UDINT;                   // +1 per cycle with every setpoint sample
    // diagnostics (bridge, HMI)
    eNewestAlarm : E_AlarmId;
    xAlarmError : BOOL;
    xAlarmCritical : BOOL;
    iWorstJoint : INT;
    aFollowingError : ARRAY[1..6] OF LREAL;   // [deg]
END_VAR
VAR
    fbSm : FB_PackMLStateMachine;
    fbAlarms : FB_AlarmHandler;
    fbSafety : FB_SafetyMonitor;
    fbConv : FB_Conveyor;
    fbRobot : FB_Robot;
    fbMon : FB_JointMonitor;
    fbTracker : FB_PartTracker;
    fbSeq : FB_PickSequence;
    fbVac : FB_VacuumGripper;
    aBins : ARRAY[E_Bin.TypeA..E_Bin.Quarantine] OF FB_Bin;
    fbPe1 : FB_PhotoEye;
    fbWatchdog : FB_BridgeWatchdog;
    fbJog : SMC_GroupJog2;
    eBin : E_Bin;
    i : INT;
    xAnyBinFull : BOOL;
    xSuspendedByBin : BOOL;             // the current suspension was caused by a full bin
    xComplete : BOOL;
    xAutoMode : BOOL;
    xRunBelt : BOOL;
    xJog : BOOL;
    xMotionStill : BOOL;                // pick sequence resting, robot and belt standing still
    lrSpeedFactor : LREAL;
    aFeedback : ARRAY[1..6] OF LREAL;
END_VAR
VAR CONSTANT
    REDUCED_SPEED_FACTOR : LREAL := 0.25;   // Maintenance mode and Manual with the door open
    JOG_VELOCITY : LREAL := 30;             // [deg/s] joint jog
    JOG_ACCELERATION : LREAL := 300;        // [deg/s2]
    JOG_JERK : LREAL := 3000;               // [deg/s3]
    JOG_MAX_LINEAR : LREAL := 100;          // [mm] per jog edge
    JOG_MAX_ANGULAR : LREAL := 45;          // [deg] per jog edge
    BELT_STANDSTILL : LREAL := 0.5;         // [mm/s] belt counts as stopped below this
END_VAR

eState := fbSm.eState;
eMode := fbSm.eMode;
xAutoMode := eMode <> E_PackMLMode.Manual;

fbRobot.itfAlarms := fbAlarms;
fbConv.itfAlarms := fbAlarms;
fbVac.itfAlarms := fbAlarms;
fbTracker.itfAlarms := fbAlarms;
fbSafety.itfAlarms := fbAlarms;
fbMon.itfAlarms := fbAlarms;
fbWatchdog.itfAlarms := fbAlarms;

// --- safety and alarm acknowledgement --------------------------------------------------------
fbSafety(xEStopOk := xEStopOk, xDoorClosed := xDoorClosed, eMode := eMode,
         xResetCmd := eState = E_PackMLState.Resetting OR eState = E_PackMLState.Clearing);
IF xAlarmAck OR (fbSm.xStateChanged AND (eState = E_PackMLState.Resetting OR eState = E_PackMLState.Clearing)) THEN
    fbAlarms.AcknowledgeAll();
END_IF

// --- bins --------------------------------------------------------------------------------------
xAnyBinFull := FALSE;
FOR eBin := E_Bin.TypeA TO E_Bin.Quarantine DO
    aBins[eBin](eBin := eBin,
                xFullSensor := axBinFull[eBin],
                xPlaced := fbSeq.xPlacedPulse AND fbSeq.eLastBin = eBin);
    xAnyBinFull := xAnyBinFull OR aBins[eBin].xFull;
END_FOR
IF xAnyBinFull THEN
    fbAlarms.Raise(E_AlarmId.BinFull);
ELSE
    fbAlarms.Clear(E_AlarmId.BinFull);
END_IF

// --- PackML state actions ----------------------------------------------------------------------
xComplete := FALSE;
xRunBelt := FALSE;
xJog := FALSE;
fbSeq.xRun := FALSE;
fbSeq.xAbort := FALSE;
fbSeq.xReset := FALSE;
xMotionStill := (fbSeq.eStep = E_PickStep.Idle OR fbSeq.eStep = E_PickStep.Error
                 OR fbSeq.eStep = E_PickStep.Aborted)
                AND NOT fbRobot.xMoving AND ABS(fbConv.lrActVelocity) < BELT_STANDSTILL;
CASE eState OF
    E_PackMLState.Resetting:
        fbSeq.xReset := TRUE;
        fbTracker.Clear();                        // parts on the belt are unknown after a stop
        fbRobot.Reset();
        fbVac.Reset();
        fbConv.Reset();
        xSuspendedByBin := FALSE;
        xComplete := fbSafety.xSafeToMove AND fbRobot.xReady AND fbSeq.eStep = E_PickStep.Idle
                     AND NOT fbAlarms.xCriticalActive AND NOT fbAlarms.xErrorActive;

    E_PackMLState.Starting, E_PackMLState.Unholding, E_PackMLState.Unsuspending:
        IF xAutoMode THEN
            fbSeq.xRun := TRUE;
            xRunBelt := TRUE;
            xComplete := fbSeq.eStep = E_PickStep.WaitPart AND fbConv.xAtSpeed;
        ELSE
            xComplete := fbRobot.xReady;
        END_IF

    E_PackMLState.Execute:
        xSuspendedByBin := xAnyBinFull;          // a full bin in Execute raises the suspension
        IF xAutoMode THEN
            fbSeq.xRun := TRUE;
            xRunBelt := TRUE;
        ELSE
            xJog := TRUE;
        END_IF

    E_PackMLState.Stopping, E_PackMLState.Holding, E_PackMLState.Suspending, E_PackMLState.Completing:
        xComplete := xMotionStill;

    E_PackMLState.Aborting:
        fbSeq.xAbort := TRUE;
        xComplete := NOT fbRobot.xMoving AND (fbSeq.eStep = E_PickStep.Aborted
                     OR fbSeq.eStep = E_PickStep.Idle OR fbSeq.eStep = E_PickStep.Error);

    E_PackMLState.Clearing:
        fbSeq.xReset := TRUE;
        fbRobot.Reset();
        fbVac.Reset();
        fbConv.Reset();
        xComplete := fbSafety.xSafeToMove AND fbSeq.eStep = E_PickStep.Idle
                     AND NOT fbAlarms.xCriticalActive;
END_CASE

// --- equipment ---------------------------------------------------------------------------------
IF eMode = E_PackMLMode.Maintenance OR fbSafety.xReducedSpeed THEN
    lrSpeedFactor := REDUCED_SPEED_FACTOR;
ELSE
    lrSpeedFactor := 1.0;
END_IF

fbPe1(xRaw := xPE1);
fbTracker(lrBeltPos := fbConv.lrPosition, xPE1Rising := fbPe1.xRising,
          stVision := stVision, stDecision := stDecision, xDecisionActive := xDecisionActive);
fbSeq(AxisGroup := AxisGroup, ConveyorAxis := ConveyorAxis,
      Robot := fbRobot, Gripper := fbVac, Tracker := fbTracker);
fbVac(xVacuumOk := xVacuumOk, tGripTimeout := GVL_Params.tVacuumTimeout);

fbRobot.xEnable := eState <> E_PackMLState.Stopped;
fbRobot.lrOverride := REAL_TO_LREAL(rOverride) * lrSpeedFactor;
fbRobot(AxisGroup := AxisGroup);

fbJog.Enable := xJog AND fbRobot.xReady AND fbSafety.xSafeToMove;
FOR i := 1 TO 6 DO
    fbJog.Forward[i - 1] := axJogPlus[i];
    fbJog.Backward[i - 1] := axJogMinus[i];
END_FOR
fbJog(AxisGroup := AxisGroup,
      CoordSystem := SMC_COORD_SYSTEM.ACS,
      MaxLinearDistance := JOG_MAX_LINEAR,
      MaxAngularDistance := JOG_MAX_ANGULAR,
      Velocity := JOG_VELOCITY,
      Acceleration := JOG_ACCELERATION,
      Deceleration := JOG_ACCELERATION,
      Jerk := JOG_JERK,
      VelFactor := lrSpeedFactor,
      AccFactor := 1.0,
      JerkFactor := 1.0);

fbConv(Axis := ConveyorAxis,
       xEnable := eState <> E_PackMLState.Stopped,
       lrVelocity := GVL_Params.lrBeltSpeed,
       xRun := xRunBelt AND fbSafety.xSafeToMove);

FOR i := 1 TO 6 DO
    IF xLoopback THEN
        aFeedback[i] := fbRobot.aSetAcs[i];
    ELSE
        aFeedback[i] := aJointPosFb[i];
    END_IF
END_FOR
udiSetpointSeq := udiSetpointSeq + 1;
fbMon(aSetpoint := fbRobot.aSetAcs, aFeedback := aFeedback, aTorque := aJointTorqueFb,
      udiFeedbackSeq := udiFeedbackSeq, udiSetpointSeq := udiSetpointSeq,
      udiFeedbackForSeq := udiFeedbackForSeq, xLoopback := xLoopback, xActive := fbRobot.xReady);
fbWatchdog(xHeartbeat := xHeartbeat, xEnable := NOT xLoopback AND eState <> E_PackMLState.Stopped);

// --- PackML ------------------------------------------------------------------------------------
fbAlarms();
fbSm(eCommand := eCommand,
     eModeRequest := eModeRequest,
     xStateComplete := xComplete,
     xAbortRequest := NOT fbSafety.xSafeToMove
                      OR (fbAlarms.xCriticalActive AND eState <> E_PackMLState.Resetting
                          AND eState <> E_PackMLState.Clearing),
     xStopRequest := fbAlarms.xErrorActive AND eState <> E_PackMLState.Resetting,
     xSuspendRequest := xAnyBinFull,
     xUnsuspendRequest := xSuspendedByBin AND NOT xAnyBinFull);

// --- outputs to the bridge ---------------------------------------------------------------------
aJointPosSp := fbRobot.aSetAcs;
lrBeltPos := fbConv.lrPosition;
lrBeltVel := fbConv.lrActVelocity;
xVacuumOn := fbVac.xValveOn;
stCapture := fbTracker.stCapture;
eState := fbSm.eState;
eMode := fbSm.eMode;
ePickStep := fbSeq.eStep;
eNewestAlarm := fbAlarms.eNewest;
xAlarmError := fbAlarms.xErrorActive;
xAlarmCritical := fbAlarms.xCriticalActive;
iWorstJoint := fbMon.iWorstJoint;
aFollowingError := fbMon.aFollowingError;
FOR i := 1 TO 6 DO
    CASE i OF
        1: aActAcs[i] := fbRobot.stActAcs.a.a0;
        2: aActAcs[i] := fbRobot.stActAcs.a.a1;
        3: aActAcs[i] := fbRobot.stActAcs.a.a2;
        4: aActAcs[i] := fbRobot.stActAcs.a.a3;
        5: aActAcs[i] := fbRobot.stActAcs.a.a4;
        6: aActAcs[i] := fbRobot.stActAcs.a.a5;
    END_CASE
END_FOR

// State of one alarm (for the HMI view).
METHOD AlarmState : ST_Alarm
VAR_INPUT
    eId : E_AlarmId;
END_VAR
AlarmState := fbAlarms.GetAlarm(eId);
END_METHOD

// Parts placed in all bins since the last reset of the counters.
METHOD PlacedCount : UINT
VAR
    eBin : E_Bin;
END_VAR
PlacedCount := 0;
FOR eBin := E_Bin.TypeA TO E_Bin.Quarantine DO
    PlacedCount := PlacedCount + aBins[eBin].uiCount;
END_FOR
END_METHOD

// TRUE while a robot motion command is active (for the HMI).
METHOD RobotMoving : BOOL
RobotMoving := fbRobot.xMoving;
END_METHOD

// TRUE while at least one bin reports full (for the HMI).
METHOD AnyBinFull : BOOL
AnyBinFull := xAnyBinFull;
END_METHOD

END_FUNCTION_BLOCK

// Device/Application/Framework/FB_PackMLStateMachine
(*
    FB_PackMLStateMachine
    Purpose : PackML unit state machine and mode manager (ISA-TR88.00.02).
    Inputs  : eCommand          - state command; acts once when it changes to a new value
              eModeRequest      - requested mode; accepted only in Stopped, Idle, Aborted
              xStateComplete    - the unit finished the current acting state
              xAbortRequest     - critical condition: abort from any state except Aborting/Aborted
              xStopRequest      - error condition: stop from Idle/Execute/Held/Suspended/acting states
              xSuspendRequest   - starved/blocked: Execute -> Suspending
              xUnsuspendRequest - Suspended -> Unsuspending
    Outputs : eState, eMode, xStateChanged (one cycle), tInState
    States  : the 17 PackML states; acting states leave on xStateComplete
*)
FUNCTION_BLOCK FB_PackMLStateMachine
VAR_INPUT
    eCommand : E_PackMLCommand;
    eModeRequest : E_PackMLMode := E_PackMLMode.Production;
    xStateComplete : BOOL;
    xAbortRequest : BOOL;
    xStopRequest : BOOL;
    xSuspendRequest : BOOL;
    xUnsuspendRequest : BOOL;
END_VAR
VAR_OUTPUT
    eState : E_PackMLState := E_PackMLState.Stopped;
    eMode : E_PackMLMode := E_PackMLMode.Production;
    xStateChanged : BOOL;
    tInState : TIME;
END_VAR
VAR
    eLastCommand : E_PackMLCommand;
    eCmd : E_PackMLCommand;              // command acting in this cycle (None if unchanged)
    eNext : E_PackMLState;
    tEntered : TIME;
END_VAR

// A command acts once, on the cycle it changes to a new value.
IF eCommand <> eLastCommand THEN
    eCmd := eCommand;
ELSE
    eCmd := E_PackMLCommand.None;
END_IF
eLastCommand := eCommand;

eNext := eState;

// An abort condition only enters Aborting; Aborting and Aborted are then handled by the state
// CASE below, so a condition that is still present (E-stop held) cannot block Aborting -> Aborted.
IF (xAbortRequest OR eCmd = E_PackMLCommand.Abort)
   AND eState <> E_PackMLState.Aborting AND eState <> E_PackMLState.Aborted THEN
    eNext := E_PackMLState.Aborting;
ELSIF (xStopRequest OR eCmd = E_PackMLCommand.Stop)
      AND eState <> E_PackMLState.Stopped AND eState <> E_PackMLState.Stopping
      AND eState <> E_PackMLState.Aborting AND eState <> E_PackMLState.Aborted
      AND eState <> E_PackMLState.Clearing THEN
    eNext := E_PackMLState.Stopping;
ELSE
    CASE eState OF
        E_PackMLState.Stopped:
            IF eCmd = E_PackMLCommand.Reset THEN eNext := E_PackMLState.Resetting; END_IF
        E_PackMLState.Resetting:
            IF xStateComplete THEN eNext := E_PackMLState.Idle; END_IF
        E_PackMLState.Idle:
            IF eCmd = E_PackMLCommand.Start THEN eNext := E_PackMLState.Starting; END_IF
        E_PackMLState.Starting:
            IF xStateComplete THEN eNext := E_PackMLState.Execute; END_IF
        E_PackMLState.Execute:
            // Producing state: it never ends on xStateComplete, only on commands/requests.
            IF eCmd = E_PackMLCommand.Hold THEN
                eNext := E_PackMLState.Holding;
            ELSIF eCmd = E_PackMLCommand.Suspend OR xSuspendRequest THEN
                eNext := E_PackMLState.Suspending;
            ELSIF eCmd = E_PackMLCommand.Complete THEN
                eNext := E_PackMLState.Completing;
            END_IF
        E_PackMLState.Holding:
            IF xStateComplete THEN eNext := E_PackMLState.Held; END_IF
        E_PackMLState.Held:
            IF eCmd = E_PackMLCommand.Unhold THEN eNext := E_PackMLState.Unholding; END_IF
        E_PackMLState.Unholding:
            IF xStateComplete THEN eNext := E_PackMLState.Execute; END_IF
        E_PackMLState.Suspending:
            IF xStateComplete THEN eNext := E_PackMLState.Suspended; END_IF
        E_PackMLState.Suspended:
            IF eCmd = E_PackMLCommand.Unsuspend OR xUnsuspendRequest THEN
                eNext := E_PackMLState.Unsuspending;
            ELSIF eCmd = E_PackMLCommand.Hold THEN
                eNext := E_PackMLState.Holding;
            END_IF
        E_PackMLState.Unsuspending:
            IF xStateComplete THEN eNext := E_PackMLState.Execute; END_IF
        E_PackMLState.Completing:
            IF xStateComplete THEN eNext := E_PackMLState.Complete; END_IF
        E_PackMLState.Complete:
            IF eCmd = E_PackMLCommand.Reset THEN eNext := E_PackMLState.Resetting; END_IF
        E_PackMLState.Stopping:
            IF xStateComplete THEN eNext := E_PackMLState.Stopped; END_IF
        E_PackMLState.Aborting:
            IF xStateComplete THEN eNext := E_PackMLState.Aborted; END_IF
        E_PackMLState.Aborted:
            IF eCmd = E_PackMLCommand.Clear THEN eNext := E_PackMLState.Clearing; END_IF
        E_PackMLState.Clearing:
            IF xStateComplete THEN eNext := E_PackMLState.Stopped; END_IF
    ELSE
        eNext := E_PackMLState.Stopped;
    END_CASE
END_IF

xStateChanged := eNext <> eState;
IF xStateChanged THEN
    eState := eNext;
    tEntered := TIME();
END_IF
tInState := TIME() - tEntered;

// Mode changes only in a resting state where no motion is commanded.
IF eModeRequest <> eMode AND (eState = E_PackMLState.Stopped OR eState = E_PackMLState.Idle
                              OR eState = E_PackMLState.Aborted) THEN
    eMode := eModeRequest;
END_IF

END_FUNCTION_BLOCK

// Device/Application/Framework/FB_AlarmHandler
(*
    FB_AlarmHandler
    Purpose : Latching alarm list (ISA-18.2 style): an alarm needs both its condition gone
              (Clear) and an acknowledgement before it leaves the list.
    Methods : Raise(eId), Clear(eId) (I_AlarmSink), AcknowledgeAll(), GetAlarm(eId)
    Outputs : xCriticalActive / xErrorActive / xWarningActive - an alarm of that class is
              active OR unacknowledged; uiActiveCount - conditions currently active;
              eNewest - last raised alarm
    Call    : the FB body once per cycle after the Raise/Clear calls of that cycle
*)
FUNCTION_BLOCK FB_AlarmHandler IMPLEMENTS I_AlarmSink
VAR_OUTPUT
    xCriticalActive : BOOL;
    xErrorActive : BOOL;
    xWarningActive : BOOL;
    uiActiveCount : UINT;
    eNewest : E_AlarmId;
END_VAR
VAR
    aAlarms : ARRAY[E_AlarmId.None..E_AlarmId.QueueOverflow] OF ST_Alarm;
    eId : E_AlarmId;
END_VAR

xCriticalActive := FALSE;
xErrorActive := FALSE;
xWarningActive := FALSE;
uiActiveCount := 0;
FOR eId := E_AlarmId.EStop TO E_AlarmId.QueueOverflow DO
    IF aAlarms[eId].xActive THEN
        uiActiveCount := uiActiveCount + 1;
    END_IF
    IF aAlarms[eId].xActive OR NOT aAlarms[eId].xAcked THEN
        CASE GVL_AlarmDefs.aDefs[eId].eClass OF
            E_AlarmClass.Critical: xCriticalActive := TRUE;
            E_AlarmClass.Error: xErrorActive := TRUE;
            E_AlarmClass.Warning: xWarningActive := TRUE;
        END_CASE
    END_IF
END_FOR

METHOD Raise
VAR_INPUT
    eId : E_AlarmId;
END_VAR
IF eId = E_AlarmId.None OR aAlarms[eId].xActive THEN
    RETURN;
END_IF
aAlarms[eId].eClass := GVL_AlarmDefs.aDefs[eId].eClass;
aAlarms[eId].xActive := TRUE;
aAlarms[eId].xAcked := FALSE;
aAlarms[eId].tRaised := TIME();
eNewest := eId;
END_METHOD

METHOD Clear
VAR_INPUT
    eId : E_AlarmId;
END_VAR
aAlarms[eId].xActive := FALSE;
END_METHOD

// Acknowledge every alarm. Active alarms stay listed until their condition clears.
METHOD AcknowledgeAll
VAR
    eId : E_AlarmId;
END_VAR
FOR eId := E_AlarmId.EStop TO E_AlarmId.QueueOverflow DO
    aAlarms[eId].xAcked := TRUE;
END_FOR
END_METHOD

METHOD GetAlarm : ST_Alarm
VAR_INPUT
    eId : E_AlarmId;
END_VAR
GetAlarm := aAlarms[eId];
END_METHOD

METHOD RaiseEvent
VAR_INPUT
    eId : E_AlarmId;
END_VAR
IF eId = E_AlarmId.None THEN
    RETURN;
END_IF
aAlarms[eId].eClass := GVL_AlarmDefs.aDefs[eId].eClass;
aAlarms[eId].xActive := FALSE;
aAlarms[eId].xAcked := FALSE;
aAlarms[eId].tRaised := TIME();
eNewest := eId;
END_METHOD

END_FUNCTION_BLOCK

// Device/Application/Interfaces/I_AlarmSink
// Anything that can receive alarms (implemented by FB_AlarmHandler).
INTERFACE I_AlarmSink

// Raise an alarm; raising an already active alarm has no effect.
METHOD Raise
VAR_INPUT
    eId : E_AlarmId;
END_VAR
END_METHOD

// The alarm condition has gone; the alarm stays listed until acknowledged.
METHOD Clear
VAR_INPUT
    eId : E_AlarmId;
END_VAR
END_METHOD

// One-shot event (no lasting condition): listed unacknowledged, never active; raised again on
// every occurrence.
METHOD RaiseEvent
VAR_INPUT
    eId : E_AlarmId;
END_VAR
END_METHOD

END_INTERFACE

// Device/Application/Equipment/FB_SafetyMonitor
(*
    FB_SafetyMonitor
    Purpose : Modelled safety logic (not certified): E-stop latch and safety door per mode.
    Inputs  : xEStopOk (TRUE = not pressed), xDoorClosed, eMode, xResetCmd, itfAlarms
    Outputs : xSafeToMove - motion allowed; xReducedSpeed - only reduced speed allowed
    Rules   : E-stop latches until xEStopOk AND xResetCmd. Door open in Production or
              Maintenance -> not safe (DoorOpen). Door open in Manual -> safe, reduced speed.
    Alarms  : EStop, DoorOpen
*)
FUNCTION_BLOCK FB_SafetyMonitor
VAR_INPUT
    xEStopOk : BOOL := TRUE;
    xDoorClosed : BOOL := TRUE;
    eMode : E_PackMLMode := E_PackMLMode.Production;
    xResetCmd : BOOL;
    itfAlarms : I_AlarmSink;
END_VAR
VAR_OUTPUT
    xSafeToMove : BOOL;
    xReducedSpeed : BOOL;
END_VAR
VAR
    xEStopLatched : BOOL;
    xDoorFault : BOOL;
END_VAR

IF NOT xEStopOk THEN
    xEStopLatched := TRUE;
ELSIF xResetCmd THEN
    xEStopLatched := FALSE;
END_IF

xDoorFault := NOT xDoorClosed AND eMode <> E_PackMLMode.Manual;
xSafeToMove := NOT xEStopLatched AND NOT xDoorFault;
xReducedSpeed := NOT xDoorClosed AND eMode = E_PackMLMode.Manual;

IF itfAlarms <> 0 THEN
    IF xEStopLatched THEN
        itfAlarms.Raise(E_AlarmId.EStop);
    ELSE
        itfAlarms.Clear(E_AlarmId.EStop);
    END_IF
    IF xDoorFault THEN
        itfAlarms.Raise(E_AlarmId.DoorOpen);
    ELSE
        itfAlarms.Clear(E_AlarmId.DoorOpen);
    END_IF
END_IF

END_FUNCTION_BLOCK

// Device/Application/Equipment/FB_Conveyor
(*
    FB_Conveyor
    Purpose : Conveyor belt on a SoftMotion axis: power, run at a velocity, halt, read back.
    In/Out  : Axis - the conveyor axis (Axis_Conveyor)
    Inputs  : xEnable - power; lrVelocity - belt speed [mm/s]; xRun - move (FALSE = halt)
    Outputs : xPowered, xAtSpeed, lrPosition [mm], lrActVelocity [mm/s]
    Alarms  : ConveyorError
*)
FUNCTION_BLOCK FB_Conveyor IMPLEMENTS I_Equipment
VAR_IN_OUT
    Axis : AXIS_REF_SM3;
END_VAR
VAR_INPUT
    xEnable : BOOL;
    lrVelocity : LREAL;
    xRun : BOOL;
    itfAlarms : I_AlarmSink;
END_VAR
VAR_OUTPUT
    xPowered : BOOL;
    xAtSpeed : BOOL;
    lrPosition : LREAL;
    lrActVelocity : LREAL;
END_VAR
VAR
    fbPower : MC_Power;
    fbMove : MC_MoveVelocity;
    fbHalt : MC_Halt;
    fbReset : MC_Reset;
    fbReadPos : MC_ReadActualPosition;
    fbReadVel : MC_ReadActualVelocity;
    lrLastVelocity : LREAL;
    xRestart : BOOL;
    xResetRequest : BOOL;
    eError : E_AlarmId;
END_VAR
VAR CONSTANT
    ACCELERATION : LREAL := 1000;      // [mm/s2]
    JERK : LREAL := 10000;             // [mm/s3]
END_VAR

fbPower(Axis := Axis, Enable := xEnable, bRegulatorOn := xEnable, bDriveStart := xEnable);
xPowered := fbPower.Status;

// A changed velocity needs a new rising edge on Execute: drop it for one cycle.
xRestart := xRun AND lrVelocity <> lrLastVelocity;
lrLastVelocity := lrVelocity;
fbMove(Axis := Axis,
       Execute := xRun AND xPowered AND NOT xRestart AND eError = E_AlarmId.None,
       Velocity := ABS(lrVelocity),
       Acceleration := ACCELERATION,
       Deceleration := ACCELERATION,
       Jerk := JERK,
       Direction := MC_Direction.positive);
fbHalt(Axis := Axis, Execute := NOT xRun AND xPowered, Deceleration := ACCELERATION, Jerk := JERK);
xAtSpeed := fbMove.InVelocity;

fbReadPos(Axis := Axis, Enable := TRUE);
fbReadVel(Axis := Axis, Enable := TRUE);
lrPosition := fbReadPos.Position;
lrActVelocity := fbReadVel.Velocity;

IF (fbPower.Error OR fbMove.Error OR fbHalt.Error) AND eError = E_AlarmId.None THEN
    eError := E_AlarmId.ConveyorError;
    IF itfAlarms <> 0 THEN
        itfAlarms.Raise(eError);
    END_IF
END_IF

fbReset(Axis := Axis, Execute := xResetRequest);
IF xResetRequest AND (fbReset.Done OR fbReset.Error) THEN
    xResetRequest := FALSE;
    IF fbReset.Done THEN
        IF itfAlarms <> 0 AND eError <> E_AlarmId.None THEN
            itfAlarms.Clear(eError);
        END_IF
        eError := E_AlarmId.None;
    END_IF
END_IF

// Requests an axis reset (done in the next FB calls). Returns TRUE when already error-free.
METHOD Reset : BOOL
IF eError <> E_AlarmId.None THEN
    xResetRequest := TRUE;
END_IF
Reset := eError = E_AlarmId.None;
END_METHOD

PROPERTY HasError : BOOL
GET
HasError := eError <> E_AlarmId.None;
END_GET
END_PROPERTY

PROPERTY ErrorId : E_AlarmId
GET
ErrorId := eError;
END_GET
END_PROPERTY

END_FUNCTION_BLOCK

// Device/Application/Interfaces/I_Equipment
// Common contract of every equipment module.
INTERFACE I_Equipment

// Clear the module's latched error. Returns TRUE when the module is error-free.
METHOD Reset : BOOL
END_METHOD

PROPERTY HasError : BOOL
GET
END_GET
END_PROPERTY

PROPERTY ErrorId : E_AlarmId
GET
END_GET
END_PROPERTY

END_INTERFACE

// Device/Application/Equipment/FB_Robot
(*
    FB_Robot
    Purpose : The 6-axis robot (SoftMotion axis group) behind a PLCopen-style command interface.
    In/Out  : AxisGroup - AxisGroup_Robot
    Inputs  : xEnable - power and enable the group
              eCmd + stTarget - command, started by a rising edge of xExecute
              lrOverride - speed override ]0, 1] for all movements
    Outputs : xReady (enabled, no error), xBusy / xDone / xError of the running command,
              eSmcError, xMoving, stActAcs, stActMcs, aSetAcs[1..6] (joint setpoints, deg)
    Alarms  : AxisGroupError
    Lag     : SoftMotion's own TCP lag check compares the virtual drives' actual position, which
              trails the setpoint by one task cycle by design; its default (1 mm) trips at speed
              with Windows task jitter. MAX_TCP_LAG covers that; the real following error of the
              servo motors is supervised by FB_JointMonitor against the twin's feedback.
    Reset   : MC_GroupReset answers "no error to reset" when the group already left ErrorStop;
              that is a successful reset (otherwise the fault, and Clearing, would never end).
              The group is enabled only while it is disabled: re-enabling a group that a reset
              left enabled is an error of MC_GroupEnable.
    Note    : call once per cycle in the SoftMotion bus cycle task.
*)
FUNCTION_BLOCK FB_Robot IMPLEMENTS I_Equipment
VAR_IN_OUT
    AxisGroup : AXIS_GROUP_REF_SM3;
END_VAR
VAR_INPUT
    xEnable : BOOL;
    eCmd : E_RobotCmd;
    stTarget : SMC_POS_REF;
    xExecute : BOOL;
    lrOverride : LREAL := 1.0;
    itfAlarms : I_AlarmSink;
END_VAR
VAR_OUTPUT
    xReady : BOOL;
    xBusy : BOOL;
    xDone : BOOL;
    xError : BOOL;
    eSmcError : SMC_ERROR;
    xMoving : BOOL;
    stActAcs : SMC_POS_REF;
    stActMcs : SMC_POS_REF;
    aSetAcs : ARRAY[1..6] OF LREAL;
END_VAR
VAR CONSTANT
    MIN_OVERRIDE : LREAL := 0.01;
    STOP_DECELERATION : LREAL := 5000;     // path deceleration of a controlled stop [mm/s2]
    STOP_JERK : LREAL := 100000;           // path jerk of a controlled stop [mm/s3]
    MAX_TCP_LAG : LREAL := 10;             // SoftMotion TCP lag tolerance [mm]
    MAX_ORIENTATION_LAG : LREAL := 2;      // [deg]
    MAX_AXIS_LAG : LREAL := 2;             // per joint [deg]
END_VAR
VAR
    fbPower : SMC_GroupPower;
    fbEnable : MC_GroupEnable;
    fbReset : MC_GroupReset;
    fbStop : MC_GroupStop := (Deceleration := STOP_DECELERATION, Jerk := STOP_JERK);
    fbOverride : MC_GroupSetOverride;
    fbPtp : MC_MoveDirectAbsolute := (CoordSystem := SMC_COORD_SYSTEM.ACS);
    fbLin : MC_MoveLinearAbsolute;
    fbReadAcs : MC_GroupReadActualPosition := (Enable := TRUE, CoordSystem := SMC_COORD_SYSTEM.ACS);
    fbReadMcs : MC_GroupReadActualPosition := (Enable := TRUE, CoordSystem := SMC_COORD_SYSTEM.MCS);
    fbReadSet : SMC_GroupReadSetPosition := (Enable := TRUE, CoordSystem := SMC_COORD_SYSTEM.ACS);
    fbStatus : MC_GroupReadStatus := (Enable := TRUE);
    fbPathTol : SMC_GroupSetPathTolerance := (MaxPositionLag := MAX_TCP_LAG,
                                              MaxOrientationLag := MAX_ORIENTATION_LAG);
    rtExecute : R_TRIG;
    eActive : E_RobotCmd;
    xResetRequest : BOOL;
    xFault : BOOL;
    lrOverrideLimited : LREAL;
    xEnabled : BOOL;                       // powered and enabled, not in error
END_VAR

rtExecute(CLK := xExecute);
IF rtExecute.Q THEN
    eActive := eCmd;
ELSIF NOT xExecute THEN
    eActive := E_RobotCmd.None;
END_IF
IF eActive = E_RobotCmd.Reset THEN
    xResetRequest := TRUE;
END_IF

fbStatus(AxisGroup := AxisGroup);
fbPower(AxisGroup := AxisGroup, Enable := xEnable, bRegulatorOn := xEnable, bDriveStart := xEnable);
fbEnable(AxisGroup := AxisGroup,
         Execute := fbPower.Status AND NOT xResetRequest
                    AND (fbStatus.GroupDisabled OR fbEnable.Busy OR fbEnable.Done));
xEnabled := fbPower.Status AND fbStatus.Valid AND NOT fbStatus.GroupDisabled
            AND NOT fbStatus.GroupErrorStop;
fbPathTol.MaxAxisLag.a0 := MAX_AXIS_LAG;
fbPathTol.MaxAxisLag.a1 := MAX_AXIS_LAG;
fbPathTol.MaxAxisLag.a2 := MAX_AXIS_LAG;
fbPathTol.MaxAxisLag.a3 := MAX_AXIS_LAG;
fbPathTol.MaxAxisLag.a4 := MAX_AXIS_LAG;
fbPathTol.MaxAxisLag.a5 := MAX_AXIS_LAG;
fbPathTol(AxisGroup := AxisGroup, Execute := xEnabled);   // again after every enable

lrOverrideLimited := LIMIT(MIN_OVERRIDE, lrOverride, 1.0);
fbOverride(AxisGroup := AxisGroup,
           Enable := xEnabled AND NOT fbStatus.GroupStopping,
           VelFactor := lrOverrideLimited,
           PathVelFactor := lrOverrideLimited);

fbPtp.Position := stTarget;
fbPtp.VelFactor := GVL_Params.lrPtpVelFactor;
IF eActive = E_RobotCmd.MovePtpMcs THEN
    fbPtp.CoordSystem := SMC_COORD_SYSTEM.MCS;
ELSE
    fbPtp.CoordSystem := SMC_COORD_SYSTEM.ACS;
END_IF
fbPtp(AxisGroup := AxisGroup, Execute := eActive = E_RobotCmd.MovePtpAcs OR eActive = E_RobotCmd.MovePtpMcs);

fbLin.Position := stTarget;
fbLin.Velocity := GVL_Params.lrLinVelocity;
fbLin.Acceleration := GVL_Params.lrLinAccel;
fbLin.Deceleration := GVL_Params.lrLinAccel;
fbLin.Jerk := GVL_Params.lrLinJerk;
IF eActive = E_RobotCmd.MoveLinPcs1 THEN
    fbLin.CoordSystem := SMC_COORD_SYSTEM.PCS_1;
ELSE
    fbLin.CoordSystem := SMC_COORD_SYSTEM.MCS;
END_IF
fbLin(AxisGroup := AxisGroup, Execute := eActive = E_RobotCmd.MoveLinMcs OR eActive = E_RobotCmd.MoveLinPcs1);

fbStop(AxisGroup := AxisGroup, Execute := eActive = E_RobotCmd.Stop);
fbReset(AxisGroup := AxisGroup, Execute := xResetRequest);
IF xResetRequest AND (fbReset.Done OR fbReset.Error) THEN
    xResetRequest := FALSE;
    IF fbReset.Done OR NOT fbStatus.GroupErrorStop THEN
        IF xFault AND itfAlarms <> 0 THEN
            itfAlarms.Clear(E_AlarmId.AxisGroupError);
        END_IF
        xFault := FALSE;
        eSmcError := SMC_ERROR.SMC_NO_ERROR;
    END_IF
    fbStatus(AxisGroup := AxisGroup);   // the fault check below must see the state after the reset
END_IF

fbReadAcs(AxisGroup := AxisGroup);
fbReadMcs(AxisGroup := AxisGroup);
fbReadSet(AxisGroup := AxisGroup);
stActAcs := fbReadAcs.Position;
stActMcs := fbReadMcs.Position;
aSetAcs[1] := fbReadSet.Position.a.a0;
aSetAcs[2] := fbReadSet.Position.a.a1;
aSetAcs[3] := fbReadSet.Position.a.a2;
aSetAcs[4] := fbReadSet.Position.a.a3;
aSetAcs[5] := fbReadSet.Position.a.a4;
aSetAcs[6] := fbReadSet.Position.a.a5;

CASE eActive OF
    E_RobotCmd.MovePtpAcs, E_RobotCmd.MovePtpMcs:
        xBusy := fbPtp.Busy; xDone := fbPtp.Done; xError := fbPtp.Error;
        IF fbPtp.Error THEN eSmcError := fbPtp.ErrorID; END_IF
    E_RobotCmd.MoveLinMcs, E_RobotCmd.MoveLinPcs1:
        xBusy := fbLin.Busy; xDone := fbLin.Done; xError := fbLin.Error;
        IF fbLin.Error THEN eSmcError := fbLin.ErrorID; END_IF
    E_RobotCmd.Stop:
        xBusy := fbStop.Busy; xDone := fbStop.Done; xError := fbStop.Error;
        IF fbStop.Error THEN eSmcError := fbStop.ErrorID; END_IF
    E_RobotCmd.Reset:
        xBusy := xResetRequest; xDone := NOT xResetRequest AND NOT xFault;
        xError := fbReset.Error AND fbStatus.GroupErrorStop;
ELSE
    xBusy := FALSE; xDone := FALSE; xError := FALSE;
END_CASE

IF (fbPower.Error OR fbEnable.Error OR fbStatus.GroupErrorStop OR xError) AND NOT xFault
   AND NOT xResetRequest THEN
    xFault := TRUE;
    IF eSmcError = SMC_ERROR.SMC_NO_ERROR THEN
        IF fbEnable.Error THEN eSmcError := fbEnable.ErrorID; ELSE eSmcError := fbPower.ErrorID; END_IF
    END_IF
    IF itfAlarms <> 0 THEN
        itfAlarms.Raise(E_AlarmId.AxisGroupError);
    END_IF
END_IF

xMoving := fbStatus.GroupMoving OR fbStatus.GroupStopping;
xReady := xEnabled AND NOT xFault;

// Requests an axis group reset (done in the next FB calls). Returns TRUE when error-free.
METHOD Reset : BOOL
IF xFault THEN
    xResetRequest := TRUE;
END_IF
Reset := NOT xFault;
END_METHOD

PROPERTY HasError : BOOL
GET
HasError := xFault;
END_GET
END_PROPERTY

PROPERTY ErrorId : E_AlarmId
GET
IF xFault THEN
    ErrorId := E_AlarmId.AxisGroupError;
ELSE
    ErrorId := E_AlarmId.None;
END_IF
END_GET
END_PROPERTY

END_FUNCTION_BLOCK

// Device/Application/Equipment/FB_JointMonitor
(*
    FB_JointMonitor
    Purpose : Supervises the robot joints against the feedback of the digital twin's servo
              motors: following error per joint and freshness of the feedback.
    Inputs  : aSetpoint / aFeedback [deg], aTorque [Nm], udiFeedbackSeq (changes with every new
              feedback sample), udiSetpointSeq (number of the current setpoint sample, +1 per
              cycle), udiFeedbackForSeq (setpoint sample the feedback answers), xLoopback
              (feedback := setpoint, no staleness check), xActive (supervision on), itfAlarms
    Outputs : aFollowingError [deg], iWorstJoint (1..6, 0 = none), xWarn, xFault, xStale
    Latency : the feedback travels through OPC UA and the twin (tens of ms). The last
              HISTORY_SIZE setpoints are kept, and the feedback is compared with the setpoint it
              answers, so transport delay does not count as following error. A feedback older
              than the history (a bridge hiccup) cannot be judged and counts as no error; if the
              feedback stays that old for tFeedbackTimeout it is stale.
    Debounce: a following error counts after CONFIRM_CYCLES cycles in a row. OPC UA does not
              hand a write to the task atomically: for one cycle the new positions may meet the
              old sequence number (a torn sample), which must not abort the cell.
    Limits  : GVL_Params.lrFollowErrWarn / lrFollowErrFault / tFeedbackTimeout
    Alarms  : FollowingErrorWarn, FollowingErrorFault, FeedbackStale
*)
FUNCTION_BLOCK FB_JointMonitor
VAR_INPUT
    aSetpoint : ARRAY[1..6] OF LREAL;
    aFeedback : ARRAY[1..6] OF LREAL;
    aTorque : ARRAY[1..6] OF LREAL;
    udiFeedbackSeq : UDINT;
    udiSetpointSeq : UDINT;
    udiFeedbackForSeq : UDINT;
    xLoopback : BOOL;
    xActive : BOOL;
    itfAlarms : I_AlarmSink;
END_VAR
VAR_OUTPUT
    aFollowingError : ARRAY[1..6] OF LREAL;
    iWorstJoint : INT;
    xWarn : BOOL;
    xFault : BOOL;
    xStale : BOOL;
END_VAR
VAR
    i : INT;
    lrWorst : LREAL;
    udiLastSeq : UDINT;
    tonStale : TON;
    aHistory : ARRAY[0..HISTORY_SIZE - 1, 1..6] OF LREAL;
    udiSlot : UDINT;
    xFromHistory : BOOL;
    uiWarnCycles : UINT;
    uiFaultCycles : UINT;
END_VAR
VAR CONSTANT
    HISTORY_SIZE : UDINT := 128;            // setpoint samples kept (512 ms at 4 ms)
    CONFIRM_CYCLES : UINT := 3;             // following error must persist this long (12 ms)
END_VAR

udiSlot := udiSetpointSeq MOD HISTORY_SIZE;
FOR i := 1 TO 6 DO
    aHistory[udiSlot, i] := aSetpoint[i];
END_FOR
// UDINT arithmetic: a feedback that answers a future setpoint wraps to a large age.
xFromHistory := udiSetpointSeq - udiFeedbackForSeq < HISTORY_SIZE;
udiSlot := udiFeedbackForSeq MOD HISTORY_SIZE;

lrWorst := 0;
iWorstJoint := 0;
FOR i := 1 TO 6 DO
    IF xLoopback OR NOT xFromHistory THEN
        aFollowingError[i] := 0;           // nothing to compare with: no judgement
    ELSE
        aFollowingError[i] := ABS(aHistory[udiSlot, i] - aFeedback[i]);
    END_IF
    IF aFollowingError[i] > lrWorst THEN
        lrWorst := aFollowingError[i];
        iWorstJoint := i;
    END_IF
END_FOR

IF xActive AND lrWorst > GVL_Params.lrFollowErrWarn THEN
    uiWarnCycles := MIN(uiWarnCycles + 1, CONFIRM_CYCLES);
ELSE
    uiWarnCycles := 0;
END_IF
IF xActive AND lrWorst > GVL_Params.lrFollowErrFault THEN
    uiFaultCycles := MIN(uiFaultCycles + 1, CONFIRM_CYCLES);
ELSE
    uiFaultCycles := 0;
END_IF
xWarn := uiWarnCycles >= CONFIRM_CYCLES;
xFault := uiFaultCycles >= CONFIRM_CYCLES;

// Feedback must keep arriving, and answer a setpoint still in the history, while supervised.
tonStale(IN := xActive AND NOT xLoopback AND (udiFeedbackSeq = udiLastSeq OR NOT xFromHistory),
         PT := GVL_Params.tFeedbackTimeout);
udiLastSeq := udiFeedbackSeq;
xStale := tonStale.Q;
xFault := xFault OR xStale;

IF itfAlarms <> 0 THEN
    IF xWarn THEN itfAlarms.Raise(E_AlarmId.FollowingErrorWarn); ELSE itfAlarms.Clear(E_AlarmId.FollowingErrorWarn); END_IF
    IF xFault AND NOT xStale THEN itfAlarms.Raise(E_AlarmId.FollowingErrorFault); ELSE itfAlarms.Clear(E_AlarmId.FollowingErrorFault); END_IF
    IF xStale THEN itfAlarms.Raise(E_AlarmId.FeedbackStale); ELSE itfAlarms.Clear(E_AlarmId.FeedbackStale); END_IF
END_IF

END_FUNCTION_BLOCK

// Device/Application/Process/FB_PartTracker
(*
    FB_PartTracker
    Purpose : Tracks every part from the PE1 capture until it is placed, missed or dropped.
              Applies vision and decision messages (only for known part ids, each message once),
              falls back to the rule-based decision at GVL_Params.tDecisionDeadline and marks
              parts that leave the pick window as missed.
    Inputs  : lrBeltPos [mm], xPE1Rising, stVision, stDecision, itfAlarms, xDecisionActive
    Outputs : stCapture (capture request to the vision service), udiPlaced/udiMissed/udiDropped,
              udiVisionMsgs (vision results applied)
    Methods : NextPickable, FindPart, GetRecord, SetState, CurrentX; property Count
    Belt X  : current X of a part = lrX (belt frame at capture) + (lrBeltPos - lrBeltPosAtCapture)
    Alarms  : QueueOverflow (condition: raised while full, cleared on the next successful capture);
              DecisionFallback, VisionMissing, LowConfidence, PartMissed (one-shot events)
*)
FUNCTION_BLOCK FB_PartTracker
VAR_INPUT
    lrBeltPos : LREAL;
    xPE1Rising : BOOL;
    stVision : ST_VisionMsg;
    stDecision : ST_DecisionMsg;
    itfAlarms : I_AlarmSink;
    // TRUE: an AI decision service answers (bridge); FALSE: the rule decides a part as soon as
    // vision has identified it, without waiting for the deadline and without DecisionFallback
    xDecisionActive : BOOL := TRUE;
END_VAR
VAR_OUTPUT
    stCapture : ST_CaptureMsg;
    udiPlaced : UDINT;
    udiMissed : UDINT;
    udiDropped : UDINT;
    udiVisionMsgs : UDINT;
END_VAR
VAR
    fbQueue : FB_PartQueue;
    fbTrigger : FB_CameraTrigger;
    fbIntake : FB_MessageIntake;
    stRec : ST_PartRecord;
    stNew : ST_PartRecord;
    uiIdx : UINT;
    i : UINT;
END_VAR

// 1. New part at the camera photo-eye.
fbTrigger(xPE1Rising := xPE1Rising, lrBeltPos := lrBeltPos);
stCapture := fbTrigger.stCapture;
IF fbTrigger.xNewPart THEN
    stRec := stNew;
    stRec.udiPartId := fbTrigger.udiNewPartId;
    stRec.lrBeltPosAtCapture := lrBeltPos;
    stRec.lrX := GVL_CellGeometry.PE1_X;         // until vision reports the exact position
    stRec.eState := E_PartState.Captured;
    stRec.tCaptured := TIME();
    IF fbQueue.AddRecord(stRec) = 0 THEN
        RaiseAlarm(E_AlarmId.QueueOverflow);
    ELSIF itfAlarms <> 0 THEN
        itfAlarms.Clear(E_AlarmId.QueueOverflow);
    END_IF
END_IF

// 2. Messages from the bridge (each sequence number once, known part ids only).
fbIntake(stVision := stVision, stDecision := stDecision);
IF fbIntake.xVisionNew THEN
    uiIdx := fbQueue.FindIndex(stVision.udiPartId);
    IF uiIdx > 0 THEN
        stRec := fbQueue.GetRecord(uiIdx);
        IF stRec.eState = E_PartState.Captured THEN
            stRec.xVisionValid := stVision.xValid;
            stRec.usiClass := stVision.usiClass;
            stRec.rConfidence := stVision.rConfidence;
            stRec.lrX := stVision.lrX;
            stRec.lrY := stVision.lrY;
            stRec.lrTheta := stVision.lrTheta;
            stRec.eState := E_PartState.Identified;
            fbQueue.PutRecord(uiIdx, stRec);
            udiVisionMsgs := udiVisionMsgs + 1;
            IF NOT xDecisionActive AND stRec.xVisionValid THEN
                stRec.eDecisionSource := E_DecisionSource.Fallback;
                stRec.eQuality := E_Quality.Unknown;
                Decide(uiIdx, stRec);
            END_IF
        END_IF
    END_IF
END_IF
IF fbIntake.xDecisionNew THEN
    uiIdx := fbQueue.FindIndex(stDecision.udiPartId);
    IF uiIdx > 0 THEN
        stRec := fbQueue.GetRecord(uiIdx);
        IF stRec.eState = E_PartState.Identified THEN
            stRec.eQuality := stDecision.eQuality;
            stRec.rQualityProb := stDecision.rQualityProb;
            stRec.xIdentReliable := stDecision.xIdentReliable;
            stRec.eDecisionSource := E_DecisionSource.Ai;
            Decide(uiIdx, stRec);
        END_IF
    END_IF
END_IF

// 3. Deadline fallback and parts leaving the pick window.
FOR i := 1 TO GVL_Config.MAX_PARTS DO
    stRec := fbQueue.GetRecord(i);
    IF (stRec.eState = E_PartState.Captured OR stRec.eState = E_PartState.Identified)
       AND TIME() - stRec.tCaptured >= GVL_Params.tDecisionDeadline THEN
        stRec.eDecisionSource := E_DecisionSource.Fallback;
        stRec.eQuality := E_Quality.Unknown;
        IF NOT stRec.xVisionValid THEN
            RaiseEventAlarm(E_AlarmId.VisionMissing);
        END_IF
        IF xDecisionActive THEN
            RaiseEventAlarm(E_AlarmId.DecisionFallback);
        END_IF
        Decide(i, stRec);
        stRec := fbQueue.GetRecord(i);
    END_IF
    IF (stRec.eState = E_PartState.Captured OR stRec.eState = E_PartState.Identified
        OR stRec.eState = E_PartState.Decided)
       AND CurrentX(i) > GVL_CellGeometry.PICK_WINDOW_END_X THEN
        SetState(i, E_PartState.Missed);
    END_IF
END_FOR

// Selects the bin, marks the record Decided and stores it.
METHOD PRIVATE Decide
VAR_INPUT
    uiIdx : UINT;
    stRecIn : ST_PartRecord;
END_VAR
VAR
    stOut : ST_PartRecord;
END_VAR
stOut := stRecIn;
stOut.eTargetBin := F_SelectBin(stOut, GVL_Params.rConfidenceThreshold, GVL_Params.aClassToBin);
stOut.eState := E_PartState.Decided;
IF stOut.xVisionValid AND stOut.rConfidence < GVL_Params.rConfidenceThreshold THEN
    RaiseEventAlarm(E_AlarmId.LowConfidence);
END_IF
fbQueue.PutRecord(uiIdx, stOut);
END_METHOD

METHOD PRIVATE RaiseAlarm
VAR_INPUT
    eId : E_AlarmId;
END_VAR
IF itfAlarms <> 0 THEN
    itfAlarms.Raise(eId);
END_IF
END_METHOD

// Current belt-frame X of the part in slot uiIdx [mm].
METHOD CurrentX : LREAL
VAR_INPUT
    uiIdx : UINT;
END_VAR
VAR
    stR : ST_PartRecord;
END_VAR
stR := fbQueue.GetRecord(uiIdx);
CurrentX := stR.lrX + (lrBeltPos - stR.lrBeltPosAtCapture);
END_METHOD

// The decided, identified part furthest downstream inside [lrMinX, lrMaxX] (belt frame), or 0.
METHOD NextPickable : UINT
VAR_INPUT
    lrMinX : LREAL;
    lrMaxX : LREAL;
END_VAR
VAR
    k : UINT;
    lrX : LREAL;
    lrBest : LREAL;
    stR : ST_PartRecord;
END_VAR
NextPickable := 0;
lrBest := lrMinX;
FOR k := 1 TO GVL_Config.MAX_PARTS DO
    stR := fbQueue.GetRecord(k);
    // a part vision did not see has no known class and height: it is not picked blind
    IF stR.eState = E_PartState.Decided AND stR.xVisionValid THEN
        lrX := CurrentX(k);
        IF lrX >= lrBest AND lrX <= lrMaxX THEN
            lrBest := lrX;
            NextPickable := k;
        END_IF
    END_IF
END_FOR
END_METHOD

// Slot index of the part with this id, or 0.
METHOD FindPart : UINT
VAR_INPUT
    udiPartId : UDINT;
END_VAR
FindPart := fbQueue.FindIndex(udiPartId);
END_METHOD

METHOD GetRecord : ST_PartRecord
VAR_INPUT
    uiIdx : UINT;
END_VAR
GetRecord := fbQueue.GetRecord(uiIdx);
END_METHOD

// Updates a part's state. Placed, Dropped and Missed parts are counted and their slot is freed;
// a missed part raises the PartMissed event.
METHOD SetState
VAR_INPUT
    uiIdx : UINT;
    eState : E_PartState;
END_VAR
VAR
    stR : ST_PartRecord;
END_VAR
stR := fbQueue.GetRecord(uiIdx);
IF stR.eState = E_PartState.Free THEN
    RETURN;
END_IF
CASE eState OF
    E_PartState.Placed:
        udiPlaced := udiPlaced + 1;
        fbQueue.Release(uiIdx);
    E_PartState.Dropped:
        udiDropped := udiDropped + 1;
        fbQueue.Release(uiIdx);
    E_PartState.Missed:
        udiMissed := udiMissed + 1;
        RaiseEventAlarm(E_AlarmId.PartMissed);
        fbQueue.Release(uiIdx);
ELSE
    stR.eState := eState;
    fbQueue.PutRecord(uiIdx, stR);
END_CASE
END_METHOD

PROPERTY Count : UINT
GET
Count := fbQueue.Count;
END_GET
END_PROPERTY

METHOD PRIVATE RaiseEventAlarm
VAR_INPUT
    eId : E_AlarmId;
END_VAR
IF itfAlarms <> 0 THEN
    itfAlarms.RaiseEvent(eId);
END_IF
END_METHOD

// Forget every tracked part (PackML Resetting: the parts on the belt are unknown, e.g. removed
// by hand while the cell was stopped). Part ids keep counting, so a late vision or decision
// message for a forgotten part matches nothing.
METHOD Clear
fbQueue.Clear();
END_METHOD

END_FUNCTION_BLOCK

// Device/Application/Framework/FB_PartQueue
(*
    FB_PartQueue
    Purpose : Fixed-capacity store of part records; a record with eState = Free is an empty slot.
    Methods : Add, FindIndex, Get, Put, Release; property Count
*)
FUNCTION_BLOCK FB_PartQueue
VAR
    aRecords : ARRAY[1..GVL_Config.MAX_PARTS] OF ST_PartRecord;
    stEmpty : ST_PartRecord;
END_VAR

// Stores the record in a free slot. Returns its index, or 0 when the queue is full.
METHOD AddRecord : UINT
VAR_INPUT
    stRec : ST_PartRecord;
END_VAR
VAR
    i : UINT;
END_VAR
AddRecord := 0;
FOR i := 1 TO GVL_Config.MAX_PARTS DO
    IF aRecords[i].eState = E_PartState.Free THEN
        aRecords[i] := stRec;
        AddRecord := i;
        RETURN;
    END_IF
END_FOR
END_METHOD

// Index of the record with this part id, or 0.
METHOD FindIndex : UINT
VAR_INPUT
    udiPartId : UDINT;
END_VAR
VAR
    i : UINT;
END_VAR
FindIndex := 0;
IF udiPartId = 0 THEN
    RETURN;
END_IF
FOR i := 1 TO GVL_Config.MAX_PARTS DO
    IF aRecords[i].eState <> E_PartState.Free AND aRecords[i].udiPartId = udiPartId THEN
        FindIndex := i;
        RETURN;
    END_IF
END_FOR
END_METHOD

METHOD GetRecord : ST_PartRecord
VAR_INPUT
    uiIdx : UINT;
END_VAR
IF uiIdx >= 1 AND uiIdx <= GVL_Config.MAX_PARTS THEN
    GetRecord := aRecords[uiIdx];
ELSE
    GetRecord := stEmpty;
END_IF
END_METHOD

METHOD PutRecord
VAR_INPUT
    uiIdx : UINT;
    stRec : ST_PartRecord;
END_VAR
IF uiIdx >= 1 AND uiIdx <= GVL_Config.MAX_PARTS THEN
    aRecords[uiIdx] := stRec;
END_IF
END_METHOD

METHOD Release
VAR_INPUT
    uiIdx : UINT;
END_VAR
IF uiIdx >= 1 AND uiIdx <= GVL_Config.MAX_PARTS THEN
    aRecords[uiIdx] := stEmpty;
END_IF
END_METHOD

PROPERTY Count : UINT
GET
VAR
    i : UINT;
END_VAR
Count := 0;
FOR i := 1 TO GVL_Config.MAX_PARTS DO
    IF aRecords[i].eState <> E_PartState.Free THEN
        Count := Count + 1;
    END_IF
END_FOR
END_GET
END_PROPERTY

// Empty every slot.
METHOD Clear
VAR
    i : UINT;
END_VAR
FOR i := 1 TO GVL_Config.MAX_PARTS DO
    aRecords[i] := stEmpty;
END_FOR
END_METHOD

END_FUNCTION_BLOCK

// Device/Application/Equipment/FB_CameraTrigger
(*
    FB_CameraTrigger
    Purpose : On the PE1 photo-eye edge, assigns a new part id and publishes a capture request
              (with the conveyor position) for the vision service.
    Outputs : stCapture (udiSeq increments per request), xNewPart (one cycle), udiNewPartId
*)
FUNCTION_BLOCK FB_CameraTrigger
VAR_INPUT
    xPE1Rising : BOOL;
    lrBeltPos : LREAL;
END_VAR
VAR_OUTPUT
    stCapture : ST_CaptureMsg;
    xNewPart : BOOL;
    udiNewPartId : UDINT;
END_VAR

xNewPart := xPE1Rising;
IF xPE1Rising THEN
    udiNewPartId := udiNewPartId + 1;
    stCapture.udiSeq := stCapture.udiSeq + 1;
    stCapture.udiPartId := udiNewPartId;
    stCapture.lrBeltPos := lrBeltPos;
END_IF

END_FUNCTION_BLOCK

// Device/Application/Comm/FB_MessageIntake
(*
    FB_MessageIntake
    Purpose : Detects new bridge messages by their sequence number, so a message written twice
              (or re-read) is processed only once.
    Outputs : xVisionNew, xDecisionNew - TRUE for one cycle per new message
*)
FUNCTION_BLOCK FB_MessageIntake
VAR_INPUT
    stVision : ST_VisionMsg;
    stDecision : ST_DecisionMsg;
END_VAR
VAR_OUTPUT
    xVisionNew : BOOL;
    xDecisionNew : BOOL;
END_VAR
VAR
    udiLastVisionSeq : UDINT;
    udiLastDecisionSeq : UDINT;
END_VAR

xVisionNew := stVision.udiSeq <> udiLastVisionSeq;
udiLastVisionSeq := stVision.udiSeq;
xDecisionNew := stDecision.udiSeq <> udiLastDecisionSeq;
udiLastDecisionSeq := stDecision.udiSeq;

END_FUNCTION_BLOCK

// Device/Application/Process/F_SelectBin
(*
    F_SelectBin
    Purpose : Bin selection of spec section 7.2:
              1. no valid vision, low confidence, or an AI decision saying the identification
                 is unreliable -> Quarantine
              2. quality Scrap -> Scrap, quality Rework -> Rework
              3. otherwise the type bin of the detected class
*)
FUNCTION F_SelectBin : E_Bin
VAR_INPUT
    stRec : ST_PartRecord;
    rConfThreshold : REAL;
    aClassToBin : ARRAY[0..2] OF E_Bin;
END_VAR

IF NOT stRec.xVisionValid OR stRec.rConfidence < rConfThreshold THEN
    F_SelectBin := E_Bin.Quarantine;
ELSIF stRec.eDecisionSource = E_DecisionSource.Ai AND NOT stRec.xIdentReliable THEN
    F_SelectBin := E_Bin.Quarantine;
ELSIF stRec.eQuality = E_Quality.Scrap THEN
    F_SelectBin := E_Bin.Scrap;
ELSIF stRec.eQuality = E_Quality.Rework THEN
    F_SelectBin := E_Bin.Rework;
ELSIF stRec.usiClass <= 2 THEN
    F_SelectBin := aClassToBin[stRec.usiClass];
ELSE
    F_SelectBin := E_Bin.Quarantine;
END_IF

END_FUNCTION

// Device/Application/Process/FB_PickSequence
(*
    FB_PickSequence
    Purpose : Pick-and-place cycle from the moving conveyor:
              home -> ready pose -> wait for a decided part in the pick window ->
              MC_TrackConveyorBelt (PCS_1 follows the part) -> linear approach / descend ->
              vacuum grip -> linear lift -> PTP to the target bin -> release -> retract.
    In/Out  : AxisGroup, ConveyorAxis, Robot (FB_Robot), Gripper (FB_VacuumGripper),
              Tracker (FB_PartTracker). The owner calls Robot, Gripper and Tracker each cycle.
    Inputs  : xRun - work on parts (FALSE: finish the current part, then go home and idle)
              xAbort - controlled stop now; the vacuum stays as it is (no dropped part)
              xReset - leave Error / Aborted to Idle. A part still held is placed in the
                       Quarantine bin on the next run; a scheduled part is marked missed.
    Outputs : eStep, xIdleAtHome, xBusy, udiPicked, udiPlaced, eLastBin, xPlacedPulse (one cycle)
    Errors  : every error first stops the robot (Aborting), then rests in Error.
    Window  : a pick is abandoned (part missed) if the part passes the pick window end before
              it is gripped.
    Moves   : linear only for the short tracked moves (PCS_1); PTP for long transfers, which
              avoids wrist/base singularities on Cartesian paths across the cell.
    Heights : approach, grip and lift heights follow the scheduled part's class
              (GVL_CellGeometry.PART_HEIGHTS).
*)
FUNCTION_BLOCK FB_PickSequence
VAR_IN_OUT
    AxisGroup : AXIS_GROUP_REF_SM3;
    ConveyorAxis : AXIS_REF_SM3;
    Robot : FB_Robot;
    Gripper : FB_VacuumGripper;
    Tracker : FB_PartTracker;
END_VAR
VAR_INPUT
    xRun : BOOL;
    xAbort : BOOL;
    xReset : BOOL;
END_VAR
VAR_OUTPUT
    eStep : E_PickStep;
    xIdleAtHome : BOOL;
    xBusy : BOOL;
    udiPicked : UDINT;
    udiPlaced : UDINT;
    eLastBin : E_Bin;
    xPlacedPulse : BOOL;
END_VAR
VAR
    fbTrack : MC_TrackConveyorBelt;
    tonRelease : TON;
    xTrackExec : BOOL;
    uiIdx : UINT;                       // slot of the part being handled, 0 = none
    stPart : ST_PartRecord;
    stObject : MC_COORD_REF;
    stTarget : SMC_POS_REF;
    stHeld : ST_PartRecord;
    xAtHome : BOOL;
    xFaultPending : BOOL;               // Aborting was entered because of an error
    xRecover : BOOL;                    // a held part must go to quarantine on the next run
    // robot command handshake
    iCmdPhase : INT;
    xRequested : BOOL;
    eReqCmd : E_RobotCmd;
    stReqTarget : SMC_POS_REF;
    xCmdDone : BOOL;
    xCmdError : BOOL;
    lrPartHeight : LREAL;               // grip height of the scheduled part's class [mm]
END_VAR
VAR CONSTANT
    RELEASE_TIME : TIME := T#200MS;      // vacuum off before retracting
END_VAR

xPlacedPulse := FALSE;
xCmdDone := FALSE;
xCmdError := FALSE;

// Robot command handshake: new command -> Execute FALSE -> TRUE -> wait for Done / Error.
CASE iCmdPhase OF
    1:
        Robot.eCmd := eReqCmd;
        Robot.stTarget := stReqTarget;
        Robot.xExecute := FALSE;
        iCmdPhase := 2;
    2:
        Robot.xExecute := TRUE;
        iCmdPhase := 3;
    3:
        IF Robot.xDone THEN
            Robot.xExecute := FALSE;
            iCmdPhase := 0;
            xCmdDone := TRUE;
        ELSIF Robot.xError THEN
            Robot.xExecute := FALSE;
            iCmdPhase := 0;
            xCmdError := TRUE;
        END_IF
END_CASE

fbTrack(AxisGroup := AxisGroup,
        ConveyorBelt := ConveyorAxis,
        Execute := xTrackExec,
        ConveyorBeltOrigin := GVL_CellGeometry.BELT_ORIGIN,
        InitialObjectPosition := stObject,
        CoordSystem := SMC_COORD_SYSTEM.PCS_1);

IF xAbort AND eStep <> E_PickStep.Idle AND eStep <> E_PickStep.Aborting
   AND eStep <> E_PickStep.Aborted AND eStep <> E_PickStep.Error THEN
    eStep := E_PickStep.Aborting;
    iCmdPhase := 0;
    xRequested := FALSE;
END_IF
IF xReset AND (eStep = E_PickStep.Error OR eStep = E_PickStep.Aborted) THEN
    IF Gripper.xHolding AND uiIdx > 0 THEN
        stPart.eTargetBin := E_Bin.Quarantine;       // unknown history: quarantine it
        xRecover := TRUE;
    ELSE
        Gripper.xCmdVacuum := FALSE;
        xRecover := FALSE;
        IF uiIdx > 0 THEN
            stHeld := Tracker.GetRecord(uiIdx);
            IF stHeld.eState = E_PartState.Scheduled OR stHeld.eState = E_PartState.Picked THEN
                Tracker.SetState(uiIdx, E_PartState.Missed);
            END_IF
            uiIdx := 0;
        END_IF
    END_IF
    eStep := E_PickStep.Idle;
    iCmdPhase := 0;
    xRequested := FALSE;
    xTrackExec := FALSE;
    xAtHome := FALSE;
    xFaultPending := FALSE;
    Robot.xExecute := FALSE;
END_IF

CASE eStep OF
    E_PickStep.Idle:
        IF xRun THEN
            IF xRecover THEN
                NextStep(E_PickStep.RecoverLift);   // a part is on the cup: straight up first
            ELSE
                NextStep(E_PickStep.MoveHome);
            END_IF
        END_IF

    E_PickStep.MoveHome:
        Request(E_RobotCmd.MovePtpAcs, GVL_CellGeometry.HOME_ACS);
        IF xCmdDone THEN
            xAtHome := TRUE;
            IF xRun THEN
                NextStep(E_PickStep.MoveReady);
            ELSE
                NextStep(E_PickStep.Idle);
            END_IF
        END_IF

    E_PickStep.RecoverLift:
        // after an abort the arm may stand anywhere (near the belt, a bin wall): lift vertically
        // to the ready height before any point-to-point move, whose path is not known
        stTarget := Robot.stActMcs;
        stTarget.c.Z := MAX(Robot.stActMcs.c.Z, GVL_CellGeometry.READY_POSE.Z);
        Request(E_RobotCmd.MoveLinMcs, stTarget);
        IF xCmdDone THEN
            NextStep(E_PickStep.MoveReady);
        END_IF

    E_PickStep.MoveReady:
        stTarget.c := GVL_CellGeometry.READY_POSE;
        Request(E_RobotCmd.MovePtpMcs, stTarget);
        IF xCmdDone THEN
            xAtHome := FALSE;
            IF xRecover THEN
                NextStep(E_PickStep.MoveToBin);     // the held part goes to its bin from Ready
            ELSE
                NextStep(E_PickStep.WaitPart);
            END_IF
        END_IF

    E_PickStep.WaitPart:
        IF NOT xRun THEN
            NextStep(E_PickStep.MoveHome);
        ELSE
            uiIdx := Tracker.NextPickable(GVL_CellGeometry.PE2_X,
                                          GVL_CellGeometry.PICK_WINDOW_END_X - GVL_CellGeometry.PICK_MARGIN);
            IF uiIdx > 0 THEN
                stPart := Tracker.GetRecord(uiIdx);
                lrPartHeight := GVL_CellGeometry.PART_HEIGHTS[MIN(stPart.usiClass, 2)];
                stObject.X := Tracker.CurrentX(uiIdx);
                stObject.Y := stPart.lrY;
                stObject.Z := GVL_CellGeometry.BELT_SURFACE_Z;
                stObject.A := stPart.lrTheta;
                stObject.B := 0;
                stObject.C := 0;
                Tracker.SetState(uiIdx, E_PartState.Scheduled);
                xTrackExec := FALSE;
                NextStep(E_PickStep.StartTracking);
            END_IF
        END_IF

    E_PickStep.StartTracking:
        xTrackExec := TRUE;
        IF fbTrack.Done THEN
            NextStep(E_PickStep.Approach);
        ELSIF fbTrack.Error THEN
            GoError();
        END_IF

    E_PickStep.Approach:
        Request(E_RobotCmd.MoveLinPcs1, TrackedPose(lrPartHeight + GVL_Params.lrApproachHeight));
        IF xCmdDone THEN
            NextStep(E_PickStep.Descend);
        END_IF

    E_PickStep.Descend:
        Request(E_RobotCmd.MoveLinPcs1, TrackedPose(lrPartHeight - GVL_Params.lrPickDepth));
        IF xCmdDone THEN
            NextStep(E_PickStep.Grip);
        END_IF

    E_PickStep.Grip:
        Gripper.xCmdVacuum := TRUE;
        IF Gripper.xHolding THEN
            Tracker.SetState(uiIdx, E_PartState.Picked);
            udiPicked := udiPicked + 1;
            NextStep(E_PickStep.Lift);
        ELSIF Gripper.HasError THEN
            Gripper.xCmdVacuum := FALSE;          // nothing is held
            Tracker.SetState(uiIdx, E_PartState.Dropped);
            uiIdx := 0;
            GoError();
        END_IF

    E_PickStep.Lift:
        Request(E_RobotCmd.MoveLinPcs1, TrackedPose(lrPartHeight + GVL_Params.lrApproachHeight));
        IF xCmdDone THEN
            xTrackExec := FALSE;
            NextStep(E_PickStep.MoveToBin);
        END_IF

    E_PickStep.MoveToBin:
        stTarget.c := GVL_CellGeometry.BIN_DROP[stPart.eTargetBin];
        Request(E_RobotCmd.MovePtpMcs, stTarget);
        IF xCmdDone THEN
            NextStep(E_PickStep.Release);
        END_IF

    E_PickStep.Release:
        Gripper.xCmdVacuum := FALSE;
        tonRelease(IN := TRUE, PT := RELEASE_TIME);
        IF tonRelease.Q THEN
            Tracker.SetState(uiIdx, E_PartState.Placed);
            uiIdx := 0;
            xRecover := FALSE;
            udiPlaced := udiPlaced + 1;
            eLastBin := stPart.eTargetBin;
            xPlacedPulse := TRUE;
            NextStep(E_PickStep.Retract);
        END_IF

    E_PickStep.Retract:
        stTarget.c := GVL_CellGeometry.BIN_DROP[stPart.eTargetBin];
        stTarget.c.Z := stTarget.c.Z + GVL_CellGeometry.RETRACT_HEIGHT;
        Request(E_RobotCmd.MoveLinMcs, stTarget);
        IF xCmdDone THEN
            IF xRun THEN
                NextStep(E_PickStep.MoveReady);
            ELSE
                NextStep(E_PickStep.MoveHome);
            END_IF
        END_IF

    E_PickStep.Aborting:
        Request(E_RobotCmd.Stop, stTarget);
        IF xCmdDone OR xCmdError THEN
            xTrackExec := FALSE;
            IF xFaultPending THEN
                xFaultPending := FALSE;
                NextStep(E_PickStep.Error);
            ELSE
                NextStep(E_PickStep.Aborted);
            END_IF
        END_IF

    E_PickStep.Aborted, E_PickStep.Error:
        ;   // wait for xReset
END_CASE

// The part passed the pick window end before it was gripped: give it up, do not chase it.
IF (eStep = E_PickStep.StartTracking OR eStep = E_PickStep.Approach OR eStep = E_PickStep.Descend
    OR eStep = E_PickStep.Grip) AND uiIdx > 0 AND NOT Gripper.xHolding
   AND Tracker.CurrentX(uiIdx) > GVL_CellGeometry.PICK_WINDOW_END_X THEN
    Gripper.xCmdVacuum := FALSE;
    Tracker.SetState(uiIdx, E_PartState.Missed);
    uiIdx := 0;
    xTrackExec := FALSE;
    iCmdPhase := 0;
    Robot.xExecute := FALSE;
    NextStep(E_PickStep.MoveReady);
END_IF

// A part lost while carrying it: stop the robot; the valve stays on (spec 5.4: no release outside
// a bin), Stopping / recovery decide what happens next.
IF (eStep = E_PickStep.Lift OR eStep = E_PickStep.MoveToBin) AND Gripper.HasError THEN
    Tracker.SetState(uiIdx, E_PartState.Dropped);
    uiIdx := 0;
    GoError();
END_IF
IF xCmdError AND eStep <> E_PickStep.Aborting AND eStep <> E_PickStep.Aborted
   AND eStep <> E_PickStep.Error THEN
    GoError();
END_IF

xIdleAtHome := eStep = E_PickStep.Idle AND xAtHome;
xBusy := eStep <> E_PickStep.Idle AND eStep <> E_PickStep.WaitPart
         AND eStep <> E_PickStep.Aborted AND eStep <> E_PickStep.Error;

// Requests a robot command once per step; the handshake in the body executes it.
METHOD PRIVATE Request
VAR_INPUT
    eCmd : E_RobotCmd;
    stTgt : SMC_POS_REF;
END_VAR
IF NOT xRequested AND iCmdPhase = 0 THEN
    eReqCmd := eCmd;
    stReqTarget := stTgt;
    iCmdPhase := 1;
    xRequested := TRUE;
END_IF
END_METHOD

METHOD PRIVATE NextStep
VAR_INPUT
    eNew : E_PickStep;
END_VAR
eStep := eNew;
xRequested := FALSE;
tonRelease(IN := FALSE);
END_METHOD

// Pose above the tracked part (PCS_1 origin) at height lrZ, tool pointing down.
METHOD PRIVATE TrackedPose : SMC_POS_REF
VAR_INPUT
    lrZ : LREAL;
END_VAR
TrackedPose.c.X := 0;
TrackedPose.c.Y := 0;
TrackedPose.c.Z := lrZ;
TrackedPose.c.A := GVL_CellGeometry.TOOL_DOWN_A;
TrackedPose.c.B := GVL_CellGeometry.TOOL_DOWN_B;
TrackedPose.c.C := GVL_CellGeometry.TOOL_DOWN_C;
END_METHOD

// Enter the error path: stop the robot first (Aborting), then rest in Error.
METHOD PRIVATE GoError
eStep := E_PickStep.Aborting;
xFaultPending := TRUE;
iCmdPhase := 0;
xRequested := FALSE;
END_METHOD

END_FUNCTION_BLOCK

